REGION Network 17: STATE Num:30 StChkPalletPrsntL1L2
   RUNG wire#powerrail
      Contact( #s30_StChkPalletPrsntL1L2 )
      wire#w1
      I_Contact( #sStWtResetRel )
      I_Contact( #s30_StChkPalletPrsntL1L2_T1 )
      I_Contact( #s30_StChkPalletPrsntL1L2_T2 )
      I_Contact( #s30_StChkPalletPrsntL1L2_T3 )
      I_Contact( #s30_StChkPalletPrsntL1L2_T4 )
      wire#w2
      Coil( #s30_StChkPalletPrsntL1L2 )
   END_RUNG
   RUNG wire#powerrail
      Contact( #s20_StWtForL1L2StoprsUp_T1 )
   END_RUNG wire#w1
   RUNG wire#w2
      { S7_GenerateENO := "TRUE" } Move(in := 30, out1 => #StateNo)
   END_RUNG
   // the same network as SCL:
   #s30_StChkPalletPrsntL1L2 := (#s30_StChkPalletPrsntL1L2 OR #s20_StWtForL1L2StoprsUp_T1) AND NOT #sStWtResetRel AND NOT #s30_StChkPalletPrsntL1L2_T1 AND NOT #s30_StChkPalletPrsntL1L2_T2 AND NOT #s30_StChkPalletPrsntL1L2_T3 AND NOT #s30_StChkPalletPrsntL1L2_T4;
   IF #s30_StChkPalletPrsntL1L2 THEN #StateNo := 30; END_IF;
END_REGION

REGION Network 18: Transition for STATE Num:40 StChkPalletAtTT
   RUNG wire#powerrail
      Contact( #s40_StChkPalletAtTT )
      I_Contact( #sStWtResetRel )
      Contact( #sSst )
      wire#w1
      I_Contact( #iPalletAtTT )
      Coil( #s40_StChkPalletAtTT_T1 )
   END_RUNG
   RUNG wire#w1
      I_Contact( #s40_StChkPalletAtTT_T1 )
      Contact( #ipalletPrsntAtTT )
      Coil( #s40_StChkPalletAtTT_T2 )
   END_RUNG
   // the same network as SCL:
   #_w1 := #s40_StChkPalletAtTT AND NOT #sStWtResetRel AND #sSst;
   #s40_StChkPalletAtTT_T1 := #_w1 AND NOT #iPalletAtTT;
   #s40_StChkPalletAtTT_T2 := #_w1 AND NOT #s40_StChkPalletAtTT_T1 AND #ipalletPrsntAtTT;
END_REGION

REGION Network 19: STATE Num:40 StChkPalletAtTT
   RUNG wire#powerrail
      Contact( #s40_StChkPalletAtTT )
      wire#w1
      I_Contact( #sStWtResetRel )
      I_Contact( #s40_StChkPalletAtTT_T1 )
      I_Contact( #s40_StChkPalletAtTT_T2 )
      wire#w2
      Coil( #s40_StChkPalletAtTT )
   END_RUNG
   RUNG wire#powerrail
      Contact( #s30_StChkPalletPrsntL1L2_T1 )
   END_RUNG wire#w1
   RUNG wire#w2
      { S7_GenerateENO := "TRUE" } Move(in := 40, out1 => #StateNo)
   END_RUNG
   // the same network as SCL:
   #s40_StChkPalletAtTT := (#s40_StChkPalletAtTT OR #s30_StChkPalletPrsntL1L2_T1) AND NOT #sStWtResetRel AND NOT #s40_StChkPalletAtTT_T1 AND NOT #s40_StChkPalletAtTT_T2;
   IF #s40_StChkPalletAtTT THEN #StateNo := 40; END_IF;
END_REGION

REGION Network 20: Transition for STATE Num:50 StWtLifterAtPos1
   RUNG wire#powerrail
      Contact( #s50_StWtLifterAtPos1 )
      I_Contact( #sStWtResetRel )
      Contact( #sSst )
      Contact( #iLifterAtPos1 )
      Coil( #s50_StWtLifterAtPos1_T1 )
   END_RUNG
   // the same network as SCL:
   #s50_StWtLifterAtPos1_T1 := #s50_StWtLifterAtPos1 AND NOT #sStWtResetRel AND #sSst AND #iLifterAtPos1;
END_REGION

REGION Network 21: STATE Num:50 StWtLifterAtPos1
   RUNG wire#powerrail
      Contact( #s50_StWtLifterAtPos1 )
      wire#w1
      I_Contact( #sStWtResetRel )
      I_Contact( #s50_StWtLifterAtPos1_T1 )
      wire#w2
      Coil( #s50_StWtLifterAtPos1 )
   END_RUNG
   RUNG wire#powerrail
      Contact( #s40_StChkPalletAtTT_T1 )
   END_RUNG wire#w1
   RUNG wire#powerrail
      Contact( #s100_StRunOutActive_T1 )
   END_RUNG wire#w1
   RUNG wire#w2
      { S7_GenerateENO := "TRUE" } Move(in := 50, out1 => #StateNo)
   END_RUNG
   // the same network as SCL:
   #s50_StWtLifterAtPos1 := (#s50_StWtLifterAtPos1 OR #s40_StChkPalletAtTT_T1 OR #s100_StRunOutActive_T1) AND NOT #sStWtResetRel AND NOT #s50_StWtLifterAtPos1_T1;
   IF #s50_StWtLifterAtPos1 THEN #StateNo := 50; END_IF;
END_REGION

REGION Network 22: Actions for STATE Num:50 StWtLifterAtPos1
   RUNG wire#powerrail
      Contact( #s50_StWtLifterAtPos1 )
      Coil( #qLifterGotoPos1 )
   END_RUNG
   // the same network as SCL:
   #qLifterGotoPos1 := #s50_StWtLifterAtPos1;
END_REGION

REGION Network 23: Transition for STATE Num:60 StWtL1S2DownOver
   RUNG wire#powerrail
      Contact( #s60_StWtL1S2DownOver )
      I_Contact( #sStWtResetRel )
      Contact( #sSst )
      Contact( #iL1S2DownOver )
      Coil( #s60_StWtL1S2DownOver_T1 )
   END_RUNG
   // the same network as SCL:
   #s60_StWtL1S2DownOver_T1 := #s60_StWtL1S2DownOver AND NOT #sStWtResetRel AND #sSst AND #iL1S2DownOver;
END_REGION

REGION Network 24: STATE Num:60 StWtL1S2DownOver
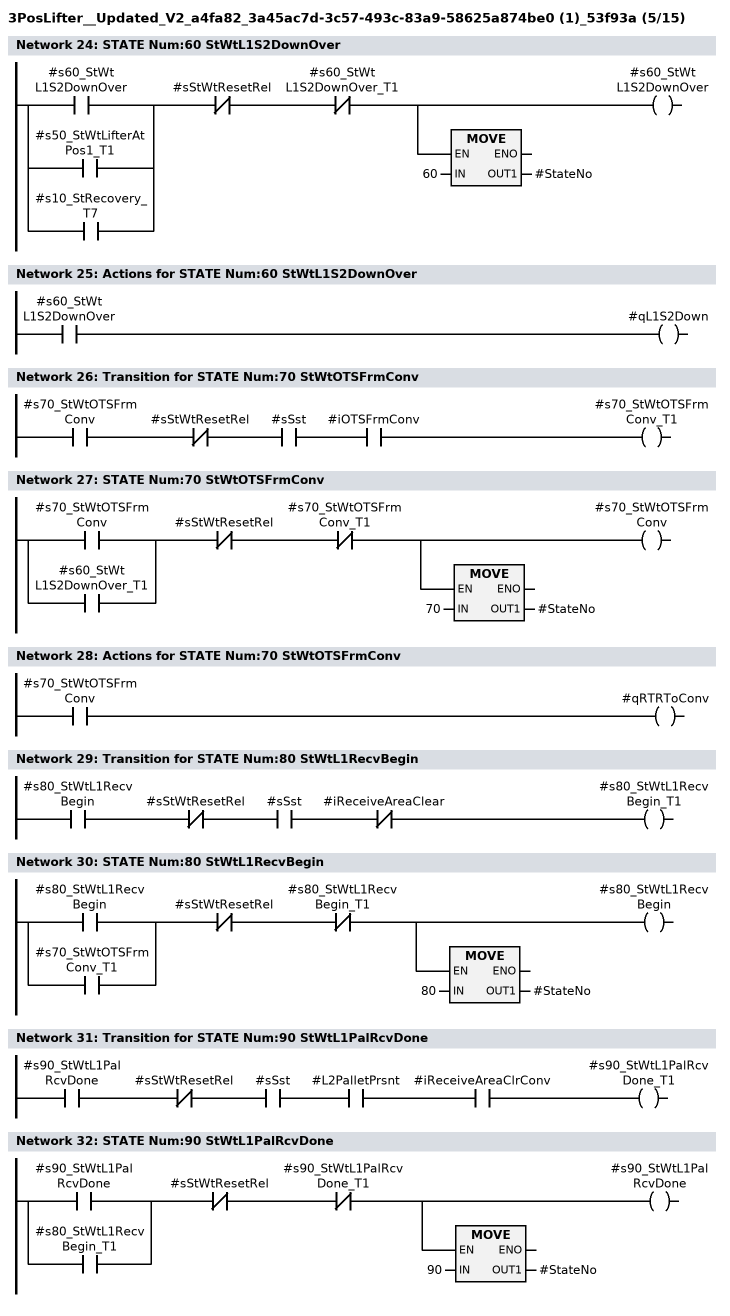
   RUNG wire#powerrail
      Contact( #s60_StWtL1S2DownOver )
      wire#w1
      I_Contact( #sStWtResetRel )
      I_Contact( #s60_StWtL1S2DownOver_T1 )
      wire#w2
      Coil( #s60_StWtL1S2DownOver )
   END_RUNG
   RUNG wire#powerrail
      Contact( #s50_StWtLifterAtPos1_T1 )
   END_RUNG wire#w1
   RUNG wire#powerrail
      Contact( #s10_StRecovery_T7 )
   END_RUNG wire#w1
   RUNG wire#w2
      { S7_GenerateENO := "TRUE" } Move(in := 60, out1 => #StateNo)
   END_RUNG
   // the same network as SCL:
   #s60_StWtL1S2DownOver := (#s60_StWtL1S2DownOver OR #s50_StWtLifterAtPos1_T1 OR #s10_StRecovery_T7) AND NOT #sStWtResetRel AND NOT #s60_StWtL1S2DownOver_T1;
   IF #s60_StWtL1S2DownOver THEN #StateNo := 60; END_IF;
END_REGION

REGION Network 25: Actions for STATE Num:60 StWtL1S2DownOver
   RUNG wire#powerrail
      Contact( #s60_StWtL1S2DownOver )
      Coil( #qL1S2Down )
   END_RUNG
   // the same network as SCL:
   #qL1S2Down := #s60_StWtL1S2DownOver;
END_REGION

REGION Network 26: Transition for STATE Num:70 StWtOTSFrmConv
   RUNG wire#powerrail
      Contact( #s70_StWtOTSFrmConv )
      I_Contact( #sStWtResetRel )
      Contact( #sSst )
      Contact( #iOTSFrmConv )
      Coil( #s70_StWtOTSFrmConv_T1 )
   END_RUNG
   // the same network as SCL:
   #s70_StWtOTSFrmConv_T1 := #s70_StWtOTSFrmConv AND NOT #sStWtResetRel AND #sSst AND #iOTSFrmConv;
END_REGION

REGION Network 27: STATE Num:70 StWtOTSFrmConv
   RUNG wire#powerrail
      Contact( #s70_StWtOTSFrmConv )
      wire#w1
      I_Contact( #sStWtResetRel )
      I_Contact( #s70_StWtOTSFrmConv_T1 )
      wire#w2
      Coil( #s70_StWtOTSFrmConv )
   END_RUNG
   RUNG wire#powerrail
      Contact( #s60_StWtL1S2DownOver_T1 )
   END_RUNG wire#w1
   RUNG wire#w2
      { S7_GenerateENO := "TRUE" } Move(in := 70, out1 => #StateNo)
   END_RUNG
   // the same network as SCL:
   #s70_StWtOTSFrmConv := (#s70_StWtOTSFrmConv OR #s60_StWtL1S2DownOver_T1) AND NOT #sStWtResetRel AND NOT #s70_StWtOTSFrmConv_T1;
   IF #s70_StWtOTSFrmConv THEN #StateNo := 70; END_IF;
END_REGION

REGION Network 28: Actions for STATE Num:70 StWtOTSFrmConv
   RUNG wire#powerrail
      Contact( #s70_StWtOTSFrmConv )
      Coil( #qRTRToConv )
   END_RUNG
   // the same network as SCL:
   #qRTRToConv := #s70_StWtOTSFrmConv;
END_REGION

REGION Network 29: Transition for STATE Num:80 StWtL1RecvBegin
   RUNG wire#powerrail
      Contact( #s80_StWtL1RecvBegin )
      I_Contact( #sStWtResetRel )
      Contact( #sSst )
      I_Contact( #iReceiveAreaClear )
      Coil( #s80_StWtL1RecvBegin_T1 )
   END_RUNG
   // the same network as SCL:
   #s80_StWtL1RecvBegin_T1 := #s80_StWtL1RecvBegin AND NOT #sStWtResetRel AND #sSst AND NOT #iReceiveAreaClear;
END_REGION

REGION Network 30: STATE Num:80 StWtL1RecvBegin
   RUNG wire#powerrail
      Contact( #s80_StWtL1RecvBegin )
      wire#w1
      I_Contact( #sStWtResetRel )
      I_Contact( #s80_StWtL1RecvBegin_T1 )
      wire#w2
      Coil( #s80_StWtL1RecvBegin )
   END_RUNG
   RUNG wire#powerrail
      Contact( #s70_StWtOTSFrmConv_T1 )
   END_RUNG wire#w1
   RUNG wire#w2
      { S7_GenerateENO := "TRUE" } Move(in := 80, out1 => #StateNo)
   END_RUNG
   // the same network as SCL:
   #s80_StWtL1RecvBegin := (#s80_StWtL1RecvBegin OR #s70_StWtOTSFrmConv_T1) AND NOT #sStWtResetRel AND NOT #s80_StWtL1RecvBegin_T1;
   IF #s80_StWtL1RecvBegin THEN #StateNo := 80; END_IF;
END_REGION

REGION Network 31: Transition for STATE Num:90 StWtL1PalRcvDone
   RUNG wire#powerrail
      Contact( #s90_StWtL1PalRcvDone )
      I_Contact( #sStWtResetRel )
      Contact( #sSst )
      Contact( #L2PalletPrsnt )
      Contact( #iReceiveAreaClrConv )
      Coil( #s90_StWtL1PalRcvDone_T1 )
   END_RUNG
   // the same network as SCL:
   #s90_StWtL1PalRcvDone_T1 := #s90_StWtL1PalRcvDone AND NOT #sStWtResetRel AND #sSst AND #L2PalletPrsnt AND #iReceiveAreaClrConv;
END_REGION

REGION Network 32: STATE Num:90 StWtL1PalRcvDone
   RUNG wire#powerrail
      Contact( #s90_StWtL1PalRcvDone )
      wire#w1
      I_Contact( #sStWtResetRel )
      I_Contact( #s90_StWtL1PalRcvDone_T1 )
      wire#w2
      Coil( #s90_StWtL1PalRcvDone )
   END_RUNG
   RUNG wire#powerrail
      Contact( #s80_StWtL1RecvBegin_T1 )
   END_RUNG wire#w1
   RUNG wire#w2
      { S7_GenerateENO := "TRUE" } Move(in := 90, out1 => #StateNo)
   END_RUNG
   // the same network as SCL:
   #s90_StWtL1PalRcvDone := (#s90_StWtL1PalRcvDone OR #s80_StWtL1RecvBegin_T1) AND NOT #sStWtResetRel AND NOT #s90_StWtL1PalRcvDone_T1;
   IF #s90_StWtL1PalRcvDone THEN #StateNo := 90; END_IF;
END_REGION

REGION Network 33: Transition for STATE Num:100 StRunOutActive
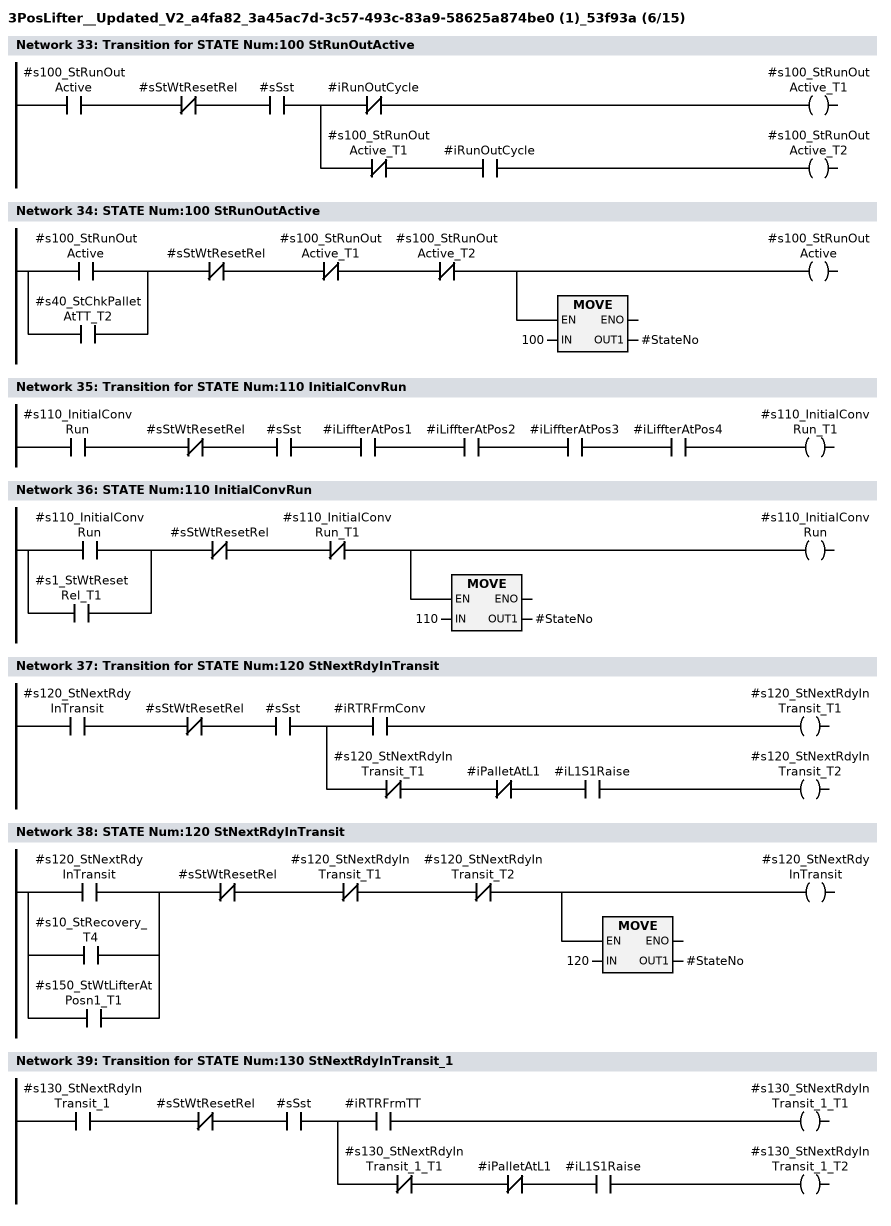
   RUNG wire#powerrail
      Contact( #s100_StRunOutActive )
      I_Contact( #sStWtResetRel )
      Contact( #sSst )
      wire#w1
      I_Contact( #iRunOutCycle )
      Coil( #s100_StRunOutActive_T1 )
   END_RUNG
   RUNG wire#w1
      I_Contact( #s100_StRunOutActive_T1 )
      Contact( #iRunOutCycle )
      Coil( #s100_StRunOutActive_T2 )
   END_RUNG
   // the same network as SCL:
   #_w1 := #s100_StRunOutActive AND NOT #sStWtResetRel AND #sSst;
   #s100_StRunOutActive_T1 := #_w1 AND NOT #iRunOutCycle;
   #s100_StRunOutActive_T2 := #_w1 AND NOT #s100_StRunOutActive_T1 AND #iRunOutCycle;
END_REGION

REGION Network 34: STATE Num:100 StRunOutActive
   RUNG wire#powerrail
      Contact( #s100_StRunOutActive )
      wire#w1
      I_Contact( #sStWtResetRel )
      I_Contact( #s100_StRunOutActive_T1 )
      I_Contact( #s100_StRunOutActive_T2 )
      wire#w2
      Coil( #s100_StRunOutActive )
   END_RUNG
   RUNG wire#powerrail
      Contact( #s40_StChkPalletAtTT_T2 )
   END_RUNG wire#w1
   RUNG wire#w2
      { S7_GenerateENO := "TRUE" } Move(in := 100, out1 => #StateNo)
   END_RUNG
   // the same network as SCL:
   #s100_StRunOutActive := (#s100_StRunOutActive OR #s40_StChkPalletAtTT_T2) AND NOT #sStWtResetRel AND NOT #s100_StRunOutActive_T1 AND NOT #s100_StRunOutActive_T2;
   IF #s100_StRunOutActive THEN #StateNo := 100; END_IF;
END_REGION

REGION Network 35: Transition for STATE Num:110 InitialConvRun
   RUNG wire#powerrail
      Contact( #s110_InitialConvRun )
      I_Contact( #sStWtResetRel )
      Contact( #sSst )
      Contact( #iLiffterAtPos1 )
      Contact( #iLiffterAtPos2 )
      Contact( #iLiffterAtPos3 )
      Contact( #iLiffterAtPos4 )
      Coil( #s110_InitialConvRun_T1 )
   END_RUNG
   // the same network as SCL:
   #s110_InitialConvRun_T1 := #s110_InitialConvRun AND NOT #sStWtResetRel AND #sSst AND #iLiffterAtPos1 AND #iLiffterAtPos2 AND #iLiffterAtPos3 AND #iLiffterAtPos4;
END_REGION

REGION Network 36: STATE Num:110 InitialConvRun
   RUNG wire#powerrail
      Contact( #s110_InitialConvRun )
      wire#w1
      I_Contact( #sStWtResetRel )
      I_Contact( #s110_InitialConvRun_T1 )
      wire#w2
      Coil( #s110_InitialConvRun )
   END_RUNG
   RUNG wire#powerrail
      Contact( #s1_StWtResetRel_T1 )
   END_RUNG wire#w1
   RUNG wire#w2
      { S7_GenerateENO := "TRUE" } Move(in := 110, out1 => #StateNo)
   END_RUNG
   // the same network as SCL:
   #s110_InitialConvRun := (#s110_InitialConvRun OR #s1_StWtResetRel_T1) AND NOT #sStWtResetRel AND NOT #s110_InitialConvRun_T1;
   IF #s110_InitialConvRun THEN #StateNo := 110; END_IF;
END_REGION

REGION Network 37: Transition for STATE Num:120 StNextRdyInTransit
   RUNG wire#powerrail
      Contact( #s120_StNextRdyInTransit )
      I_Contact( #sStWtResetRel )
      Contact( #sSst )
      wire#w1
      Contact( #iRTRFrmConv )
      Coil( #s120_StNextRdyInTransit_T1 )
   END_RUNG
   RUNG wire#w1
      I_Contact( #s120_StNextRdyInTransit_T1 )
      I_Contact( #iPalletAtL1 )
      Contact( #iL1S1Raise )
      Coil( #s120_StNextRdyInTransit_T2 )
   END_RUNG
   // the same network as SCL:
   #_w1 := #s120_StNextRdyInTransit AND NOT #sStWtResetRel AND #sSst;
   #s120_StNextRdyInTransit_T1 := #_w1 AND #iRTRFrmConv;
   #s120_StNextRdyInTransit_T2 := #_w1 AND NOT #s120_StNextRdyInTransit_T1 AND NOT #iPalletAtL1 AND #iL1S1Raise;
END_REGION

REGION Network 38: STATE Num:120 StNextRdyInTransit
   RUNG wire#powerrail
      Contact( #s120_StNextRdyInTransit )
      wire#w1
      I_Contact( #sStWtResetRel )
      I_Contact( #s120_StNextRdyInTransit_T1 )
      I_Contact( #s120_StNextRdyInTransit_T2 )
      wire#w2
      Coil( #s120_StNextRdyInTransit )
   END_RUNG
   RUNG wire#powerrail
      Contact( #s10_StRecovery_T4 )
   END_RUNG wire#w1
   RUNG wire#powerrail
      Contact( #s150_StWtLifterAtPosn1_T1 )
   END_RUNG wire#w1
   RUNG wire#w2
      { S7_GenerateENO := "TRUE" } Move(in := 120, out1 => #StateNo)
   END_RUNG
   // the same network as SCL:
   #s120_StNextRdyInTransit := (#s120_StNextRdyInTransit OR #s10_StRecovery_T4 OR #s150_StWtLifterAtPosn1_T1) AND NOT #sStWtResetRel AND NOT #s120_StNextRdyInTransit_T1 AND NOT #s120_StNextRdyInTransit_T2;
   IF #s120_StNextRdyInTransit THEN #StateNo := 120; END_IF;
END_REGION

REGION Network 39: Transition for STATE Num:130 StNextRdyInTransit_1
   RUNG wire#powerrail
      Contact( #s130_StNextRdyInTransit_1 )
      I_Contact( #sStWtResetRel )
      Contact( #sSst )
      wire#w1
      Contact( #iRTRFrmTT )
      Coil( #s130_StNextRdyInTransit_1_T1 )
   END_RUNG
   RUNG wire#w1
      I_Contact( #s130_StNextRdyInTransit_1_T1 )
      I_Contact( #iPalletAtL1 )
      Contact( #iL1S1Raise )
      Coil( #s130_StNextRdyInTransit_1_T2 )
   END_RUNG
   // the same network as SCL:
   #_w1 := #s130_StNextRdyInTransit_1 AND NOT #sStWtResetRel AND #sSst;
   #s130_StNextRdyInTransit_1_T1 := #_w1 AND #iRTRFrmTT;
   #s130_StNextRdyInTransit_1_T2 := #_w1 AND NOT #s130_StNextRdyInTransit_1_T1 AND NOT #iPalletAtL1 AND #iL1S1Raise;
END_REGION

REGION Network 40: STATE Num:130 StNextRdyInTransit_1
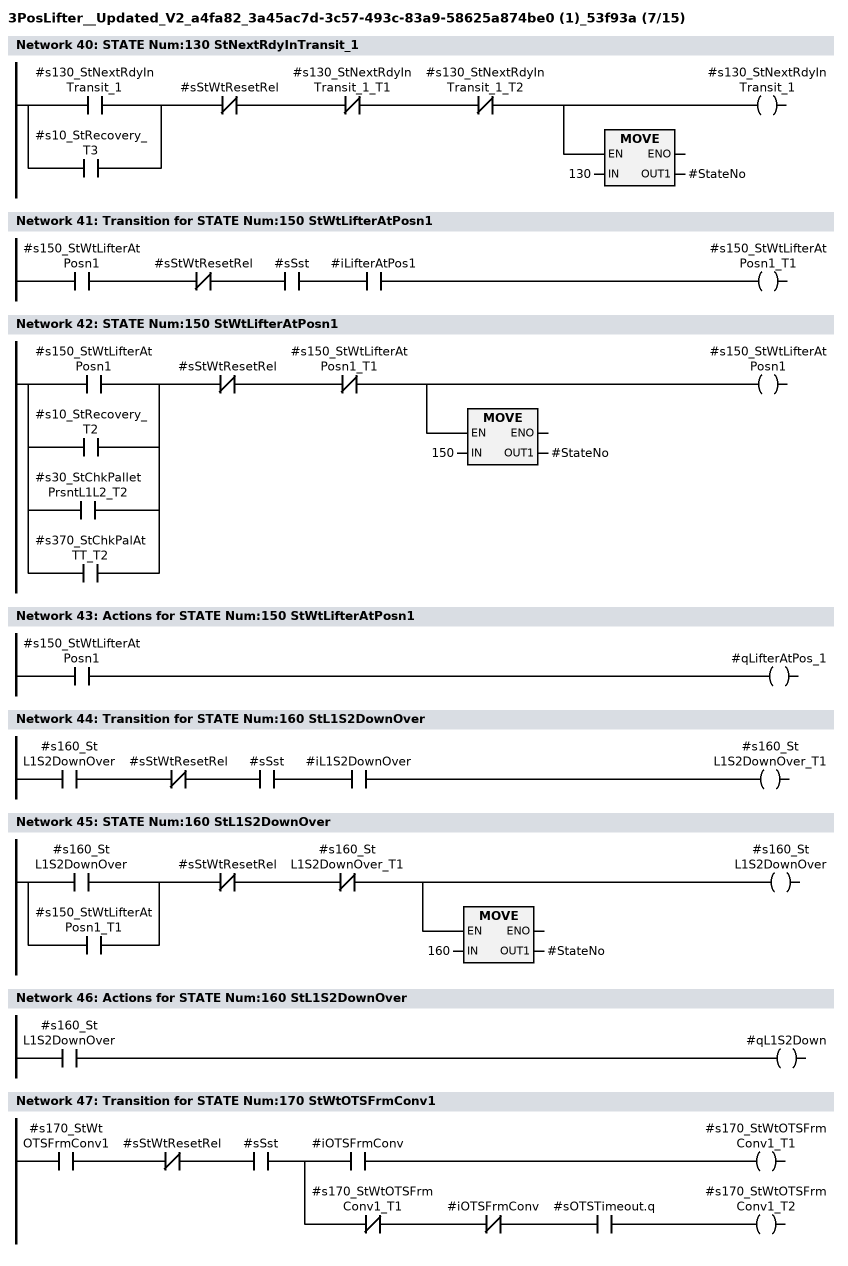
   RUNG wire#powerrail
      Contact( #s130_StNextRdyInTransit_1 )
      wire#w1
      I_Contact( #sStWtResetRel )
      I_Contact( #s130_StNextRdyInTransit_1_T1 )
      I_Contact( #s130_StNextRdyInTransit_1_T2 )
      wire#w2
      Coil( #s130_StNextRdyInTransit_1 )
   END_RUNG
   RUNG wire#powerrail
      Contact( #s10_StRecovery_T3 )
   END_RUNG wire#w1
   RUNG wire#w2
      { S7_GenerateENO := "TRUE" } Move(in := 130, out1 => #StateNo)
   END_RUNG
   // the same network as SCL:
   #s130_StNextRdyInTransit_1 := (#s130_StNextRdyInTransit_1 OR #s10_StRecovery_T3) AND NOT #sStWtResetRel AND NOT #s130_StNextRdyInTransit_1_T1 AND NOT #s130_StNextRdyInTransit_1_T2;
   IF #s130_StNextRdyInTransit_1 THEN #StateNo := 130; END_IF;
END_REGION

REGION Network 41: Transition for STATE Num:150 StWtLifterAtPosn1
   RUNG wire#powerrail
      Contact( #s150_StWtLifterAtPosn1 )
      I_Contact( #sStWtResetRel )
      Contact( #sSst )
      Contact( #iLifterAtPos1 )
      Coil( #s150_StWtLifterAtPosn1_T1 )
   END_RUNG
   // the same network as SCL:
   #s150_StWtLifterAtPosn1_T1 := #s150_StWtLifterAtPosn1 AND NOT #sStWtResetRel AND #sSst AND #iLifterAtPos1;
END_REGION

REGION Network 42: STATE Num:150 StWtLifterAtPosn1
   RUNG wire#powerrail
      Contact( #s150_StWtLifterAtPosn1 )
      wire#w1
      I_Contact( #sStWtResetRel )
      I_Contact( #s150_StWtLifterAtPosn1_T1 )
      wire#w2
      Coil( #s150_StWtLifterAtPosn1 )
   END_RUNG
   RUNG wire#powerrail
      Contact( #s10_StRecovery_T2 )
   END_RUNG wire#w1
   RUNG wire#powerrail
      Contact( #s30_StChkPalletPrsntL1L2_T2 )
   END_RUNG wire#w1
   RUNG wire#powerrail
      Contact( #s370_StChkPalAtTT_T2 )
   END_RUNG wire#w1
   RUNG wire#w2
      { S7_GenerateENO := "TRUE" } Move(in := 150, out1 => #StateNo)
   END_RUNG
   // the same network as SCL:
   #s150_StWtLifterAtPosn1 := (#s150_StWtLifterAtPosn1 OR #s10_StRecovery_T2 OR #s30_StChkPalletPrsntL1L2_T2 OR #s370_StChkPalAtTT_T2) AND NOT #sStWtResetRel AND NOT #s150_StWtLifterAtPosn1_T1;
   IF #s150_StWtLifterAtPosn1 THEN #StateNo := 150; END_IF;
END_REGION

REGION Network 43: Actions for STATE Num:150 StWtLifterAtPosn1
   RUNG wire#powerrail
      Contact( #s150_StWtLifterAtPosn1 )
      Coil( #qLifterAtPos_1 )
   END_RUNG
   // the same network as SCL:
   #qLifterAtPos_1 := #s150_StWtLifterAtPosn1;
END_REGION

REGION Network 44: Transition for STATE Num:160 StL1S2DownOver
   RUNG wire#powerrail
      Contact( #s160_StL1S2DownOver )
      I_Contact( #sStWtResetRel )
      Contact( #sSst )
      Contact( #iL1S2DownOver )
      Coil( #s160_StL1S2DownOver_T1 )
   END_RUNG
   // the same network as SCL:
   #s160_StL1S2DownOver_T1 := #s160_StL1S2DownOver AND NOT #sStWtResetRel AND #sSst AND #iL1S2DownOver;
END_REGION

REGION Network 45: STATE Num:160 StL1S2DownOver
   RUNG wire#powerrail
      Contact( #s160_StL1S2DownOver )
      wire#w1
      I_Contact( #sStWtResetRel )
      I_Contact( #s160_StL1S2DownOver_T1 )
      wire#w2
      Coil( #s160_StL1S2DownOver )
   END_RUNG
   RUNG wire#powerrail
      Contact( #s150_StWtLifterAtPosn1_T1 )
   END_RUNG wire#w1
   RUNG wire#w2
      { S7_GenerateENO := "TRUE" } Move(in := 160, out1 => #StateNo)
   END_RUNG
   // the same network as SCL:
   #s160_StL1S2DownOver := (#s160_StL1S2DownOver OR #s150_StWtLifterAtPosn1_T1) AND NOT #sStWtResetRel AND NOT #s160_StL1S2DownOver_T1;
   IF #s160_StL1S2DownOver THEN #StateNo := 160; END_IF;
END_REGION

REGION Network 46: Actions for STATE Num:160 StL1S2DownOver
   RUNG wire#powerrail
      Contact( #s160_StL1S2DownOver )
      Coil( #qL1S2Down )
   END_RUNG
   // the same network as SCL:
   #qL1S2Down := #s160_StL1S2DownOver;
END_REGION

REGION Network 47: Transition for STATE Num:170 StWtOTSFrmConv1
   RUNG wire#powerrail
      Contact( #s170_StWtOTSFrmConv1 )
      I_Contact( #sStWtResetRel )
      Contact( #sSst )
      wire#w1
      Contact( #iOTSFrmConv )
      Coil( #s170_StWtOTSFrmConv1_T1 )
   END_RUNG
   RUNG wire#w1
      I_Contact( #s170_StWtOTSFrmConv1_T1 )
      I_Contact( #iOTSFrmConv )
      Contact( #sOTSTimeout.q )
      Coil( #s170_StWtOTSFrmConv1_T2 )
   END_RUNG
   // the same network as SCL:
   #_w1 := #s170_StWtOTSFrmConv1 AND NOT #sStWtResetRel AND #sSst;
   #s170_StWtOTSFrmConv1_T1 := #_w1 AND #iOTSFrmConv;
   #s170_StWtOTSFrmConv1_T2 := #_w1 AND NOT #s170_StWtOTSFrmConv1_T1 AND NOT #iOTSFrmConv AND #sOTSTimeout.q;
END_REGION

REGION Network 48: STATE Num:170 StWtOTSFrmConv1
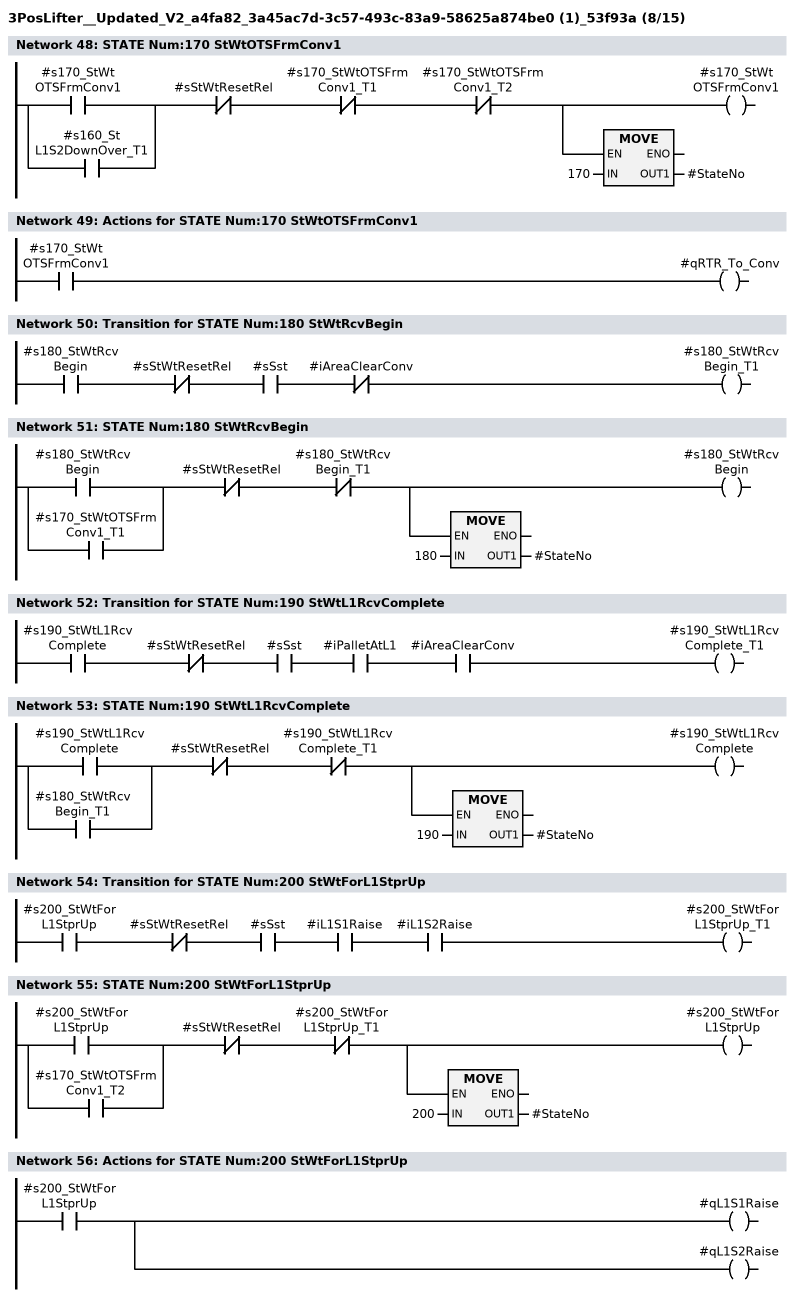
   RUNG wire#powerrail
      Contact( #s170_StWtOTSFrmConv1 )
      wire#w1
      I_Contact( #sStWtResetRel )
      I_Contact( #s170_StWtOTSFrmConv1_T1 )
      I_Contact( #s170_StWtOTSFrmConv1_T2 )
      wire#w2
      Coil( #s170_StWtOTSFrmConv1 )
   END_RUNG
   RUNG wire#powerrail
      Contact( #s160_StL1S2DownOver_T1 )
   END_RUNG wire#w1
   RUNG wire#w2
      { S7_GenerateENO := "TRUE" } Move(in := 170, out1 => #StateNo)
   END_RUNG
   // the same network as SCL:
   #s170_StWtOTSFrmConv1 := (#s170_StWtOTSFrmConv1 OR #s160_StL1S2DownOver_T1) AND NOT #sStWtResetRel AND NOT #s170_StWtOTSFrmConv1_T1 AND NOT #s170_StWtOTSFrmConv1_T2;
   IF #s170_StWtOTSFrmConv1 THEN #StateNo := 170; END_IF;
END_REGION

REGION Network 49: Actions for STATE Num:170 StWtOTSFrmConv1
   RUNG wire#powerrail
      Contact( #s170_StWtOTSFrmConv1 )
      Coil( #qRTR_To_Conv )
   END_RUNG
   // the same network as SCL:
   #qRTR_To_Conv := #s170_StWtOTSFrmConv1;
END_REGION

REGION Network 50: Transition for STATE Num:180 StWtRcvBegin
   RUNG wire#powerrail
      Contact( #s180_StWtRcvBegin )
      I_Contact( #sStWtResetRel )
      Contact( #sSst )
      I_Contact( #iAreaClearConv )
      Coil( #s180_StWtRcvBegin_T1 )
   END_RUNG
   // the same network as SCL:
   #s180_StWtRcvBegin_T1 := #s180_StWtRcvBegin AND NOT #sStWtResetRel AND #sSst AND NOT #iAreaClearConv;
END_REGION

REGION Network 51: STATE Num:180 StWtRcvBegin
   RUNG wire#powerrail
      Contact( #s180_StWtRcvBegin )
      wire#w1
      I_Contact( #sStWtResetRel )
      I_Contact( #s180_StWtRcvBegin_T1 )
      wire#w2
      Coil( #s180_StWtRcvBegin )
   END_RUNG
   RUNG wire#powerrail
      Contact( #s170_StWtOTSFrmConv1_T1 )
   END_RUNG wire#w1
   RUNG wire#w2
      { S7_GenerateENO := "TRUE" } Move(in := 180, out1 => #StateNo)
   END_RUNG
   // the same network as SCL:
   #s180_StWtRcvBegin := (#s180_StWtRcvBegin OR #s170_StWtOTSFrmConv1_T1) AND NOT #sStWtResetRel AND NOT #s180_StWtRcvBegin_T1;
   IF #s180_StWtRcvBegin THEN #StateNo := 180; END_IF;
END_REGION

REGION Network 52: Transition for STATE Num:190 StWtL1RcvComplete
   RUNG wire#powerrail
      Contact( #s190_StWtL1RcvComplete )
      I_Contact( #sStWtResetRel )
      Contact( #sSst )
      Contact( #iPalletAtL1 )
      Contact( #iAreaClearConv )
      Coil( #s190_StWtL1RcvComplete_T1 )
   END_RUNG
   // the same network as SCL:
   #s190_StWtL1RcvComplete_T1 := #s190_StWtL1RcvComplete AND NOT #sStWtResetRel AND #sSst AND #iPalletAtL1 AND #iAreaClearConv;
END_REGION

REGION Network 53: STATE Num:190 StWtL1RcvComplete
   RUNG wire#powerrail
      Contact( #s190_StWtL1RcvComplete )
      wire#w1
      I_Contact( #sStWtResetRel )
      I_Contact( #s190_StWtL1RcvComplete_T1 )
      wire#w2
      Coil( #s190_StWtL1RcvComplete )
   END_RUNG
   RUNG wire#powerrail
      Contact( #s180_StWtRcvBegin_T1 )
   END_RUNG wire#w1
   RUNG wire#w2
      { S7_GenerateENO := "TRUE" } Move(in := 190, out1 => #StateNo)
   END_RUNG
   // the same network as SCL:
   #s190_StWtL1RcvComplete := (#s190_StWtL1RcvComplete OR #s180_StWtRcvBegin_T1) AND NOT #sStWtResetRel AND NOT #s190_StWtL1RcvComplete_T1;
   IF #s190_StWtL1RcvComplete THEN #StateNo := 190; END_IF;
END_REGION

REGION Network 54: Transition for STATE Num:200 StWtForL1StprUp
   RUNG wire#powerrail
      Contact( #s200_StWtForL1StprUp )
      I_Contact( #sStWtResetRel )
      Contact( #sSst )
      Contact( #iL1S1Raise )
      Contact( #iL1S2Raise )
      Coil( #s200_StWtForL1StprUp_T1 )
   END_RUNG
   // the same network as SCL:
   #s200_StWtForL1StprUp_T1 := #s200_StWtForL1StprUp AND NOT #sStWtResetRel AND #sSst AND #iL1S1Raise AND #iL1S2Raise;
END_REGION

REGION Network 55: STATE Num:200 StWtForL1StprUp
   RUNG wire#powerrail
      Contact( #s200_StWtForL1StprUp )
      wire#w1
      I_Contact( #sStWtResetRel )
      I_Contact( #s200_StWtForL1StprUp_T1 )
      wire#w2
      Coil( #s200_StWtForL1StprUp )
   END_RUNG
   RUNG wire#powerrail
      Contact( #s170_StWtOTSFrmConv1_T2 )
   END_RUNG wire#w1
   RUNG wire#w2
      { S7_GenerateENO := "TRUE" } Move(in := 200, out1 => #StateNo)
   END_RUNG
   // the same network as SCL:
   #s200_StWtForL1StprUp := (#s200_StWtForL1StprUp OR #s170_StWtOTSFrmConv1_T2) AND NOT #sStWtResetRel AND NOT #s200_StWtForL1StprUp_T1;
   IF #s200_StWtForL1StprUp THEN #StateNo := 200; END_IF;
END_REGION

REGION Network 56: Actions for STATE Num:200 StWtForL1StprUp
   RUNG wire#powerrail
      Contact( #s200_StWtForL1StprUp )
      wire#w1
      Coil( #qL1S1Raise )
   END_RUNG
   RUNG wire#w1
      Coil( #qL1S2Raise )
   END_RUNG
   // the same network as SCL:
   #qL1S1Raise := #s200_StWtForL1StprUp;
   #qL1S2Raise := #s200_StWtForL1StprUp;
END_REGION

REGION Network 57: Transition for STATE Num:220 StWtL2S2Down
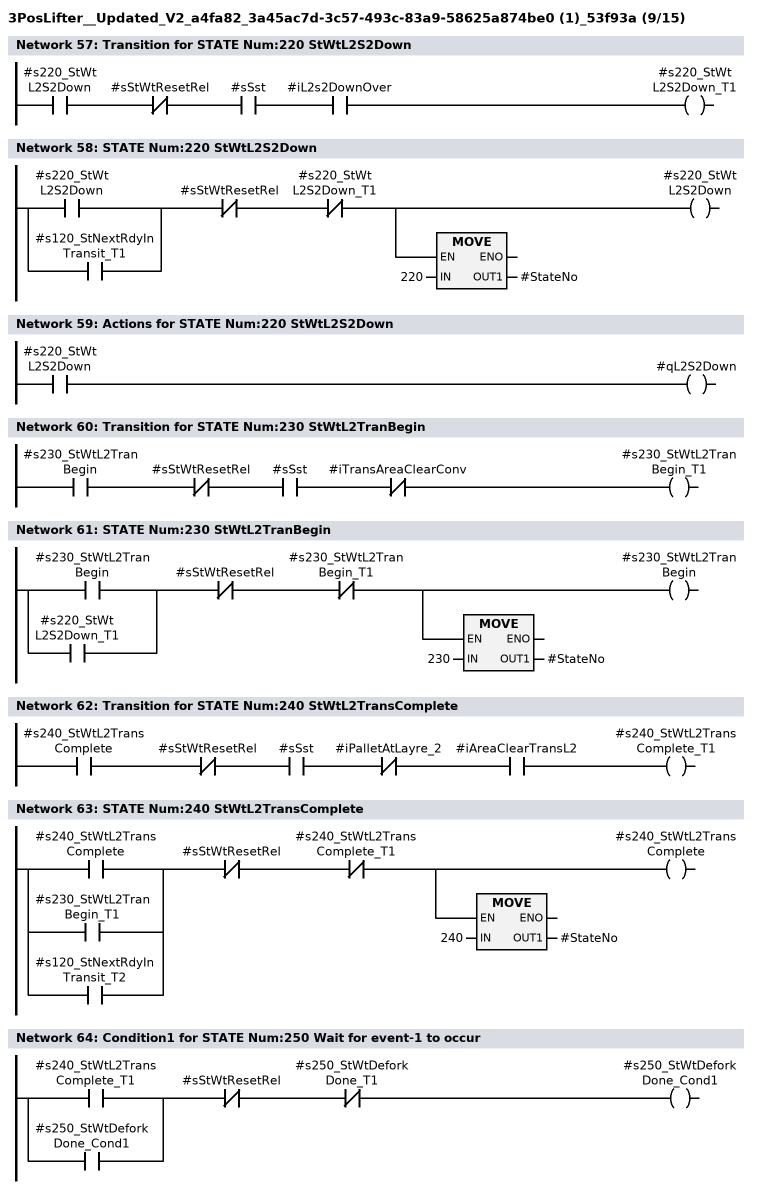
   RUNG wire#powerrail
      Contact( #s220_StWtL2S2Down )
      I_Contact( #sStWtResetRel )
      Contact( #sSst )
      Contact( #iL2s2DownOver )
      Coil( #s220_StWtL2S2Down_T1 )
   END_RUNG
   // the same network as SCL:
   #s220_StWtL2S2Down_T1 := #s220_StWtL2S2Down AND NOT #sStWtResetRel AND #sSst AND #iL2s2DownOver;
END_REGION

REGION Network 58: STATE Num:220 StWtL2S2Down
   RUNG wire#powerrail
      Contact( #s220_StWtL2S2Down )
      wire#w1
      I_Contact( #sStWtResetRel )
      I_Contact( #s220_StWtL2S2Down_T1 )
      wire#w2
      Coil( #s220_StWtL2S2Down )
   END_RUNG
   RUNG wire#powerrail
      Contact( #s120_StNextRdyInTransit_T1 )
   END_RUNG wire#w1
   RUNG wire#w2
      { S7_GenerateENO := "TRUE" } Move(in := 220, out1 => #StateNo)
   END_RUNG
   // the same network as SCL:
   #s220_StWtL2S2Down := (#s220_StWtL2S2Down OR #s120_StNextRdyInTransit_T1) AND NOT #sStWtResetRel AND NOT #s220_StWtL2S2Down_T1;
   IF #s220_StWtL2S2Down THEN #StateNo := 220; END_IF;
END_REGION

REGION Network 59: Actions for STATE Num:220 StWtL2S2Down
   RUNG wire#powerrail
      Contact( #s220_StWtL2S2Down )
      Coil( #qL2S2Down )
   END_RUNG
   // the same network as SCL:
   #qL2S2Down := #s220_StWtL2S2Down;
END_REGION

REGION Network 60: Transition for STATE Num:230 StWtL2TranBegin
   RUNG wire#powerrail
      Contact( #s230_StWtL2TranBegin )
      I_Contact( #sStWtResetRel )
      Contact( #sSst )
      I_Contact( #iTransAreaClearConv )
      Coil( #s230_StWtL2TranBegin_T1 )
   END_RUNG
   // the same network as SCL:
   #s230_StWtL2TranBegin_T1 := #s230_StWtL2TranBegin AND NOT #sStWtResetRel AND #sSst AND NOT #iTransAreaClearConv;
END_REGION

REGION Network 61: STATE Num:230 StWtL2TranBegin
   RUNG wire#powerrail
      Contact( #s230_StWtL2TranBegin )
      wire#w1
      I_Contact( #sStWtResetRel )
      I_Contact( #s230_StWtL2TranBegin_T1 )
      wire#w2
      Coil( #s230_StWtL2TranBegin )
   END_RUNG
   RUNG wire#powerrail
      Contact( #s220_StWtL2S2Down_T1 )
   END_RUNG wire#w1
   RUNG wire#w2
      { S7_GenerateENO := "TRUE" } Move(in := 230, out1 => #StateNo)
   END_RUNG
   // the same network as SCL:
   #s230_StWtL2TranBegin := (#s230_StWtL2TranBegin OR #s220_StWtL2S2Down_T1) AND NOT #sStWtResetRel AND NOT #s230_StWtL2TranBegin_T1;
   IF #s230_StWtL2TranBegin THEN #StateNo := 230; END_IF;
END_REGION

REGION Network 62: Transition for STATE Num:240 StWtL2TransComplete
   RUNG wire#powerrail
      Contact( #s240_StWtL2TransComplete )
      I_Contact( #sStWtResetRel )
      Contact( #sSst )
      I_Contact( #iPalletAtLayre_2 )
      Contact( #iAreaClearTransL2 )
      Coil( #s240_StWtL2TransComplete_T1 )
   END_RUNG
   // the same network as SCL:
   #s240_StWtL2TransComplete_T1 := #s240_StWtL2TransComplete AND NOT #sStWtResetRel AND #sSst AND NOT #iPalletAtLayre_2 AND #iAreaClearTransL2;
END_REGION

REGION Network 63: STATE Num:240 StWtL2TransComplete
   RUNG wire#powerrail
      Contact( #s240_StWtL2TransComplete )
      wire#w1
      I_Contact( #sStWtResetRel )
      I_Contact( #s240_StWtL2TransComplete_T1 )
      wire#w2
      Coil( #s240_StWtL2TransComplete )
   END_RUNG
   RUNG wire#powerrail
      Contact( #s230_StWtL2TranBegin_T1 )
   END_RUNG wire#w1
   RUNG wire#powerrail
      Contact( #s120_StNextRdyInTransit_T2 )
   END_RUNG wire#w1
   RUNG wire#w2
      { S7_GenerateENO := "TRUE" } Move(in := 240, out1 => #StateNo)
   END_RUNG
   // the same network as SCL:
   #s240_StWtL2TransComplete := (#s240_StWtL2TransComplete OR #s230_StWtL2TranBegin_T1 OR #s120_StNextRdyInTransit_T2) AND NOT #sStWtResetRel AND NOT #s240_StWtL2TransComplete_T1;
   IF #s240_StWtL2TransComplete THEN #StateNo := 240; END_IF;
END_REGION

REGION Network 64: Condition1 for STATE Num:250 Wait for event-1 to occur
   RUNG wire#powerrail
      Contact( #s240_StWtL2TransComplete_T1 )
      wire#w1
      I_Contact( #sStWtResetRel )
      I_Contact( #s250_StWtDeforkDone_T1 )
      Coil( #s250_StWtDeforkDone_Cond1 )
   END_RUNG
   RUNG wire#powerrail
      Contact( #s250_StWtDeforkDone_Cond1 )
   END_RUNG wire#w1
   // the same network as SCL:
   #s250_StWtDeforkDone_Cond1 := (#s240_StWtL2TransComplete_T1 OR #s250_StWtDeforkDone_Cond1) AND NOT #sStWtResetRel AND NOT #s250_StWtDeforkDone_T1;
END_REGION

REGION Network 65: Condition2 for STATE Num:250 Wait for event-1 to occur
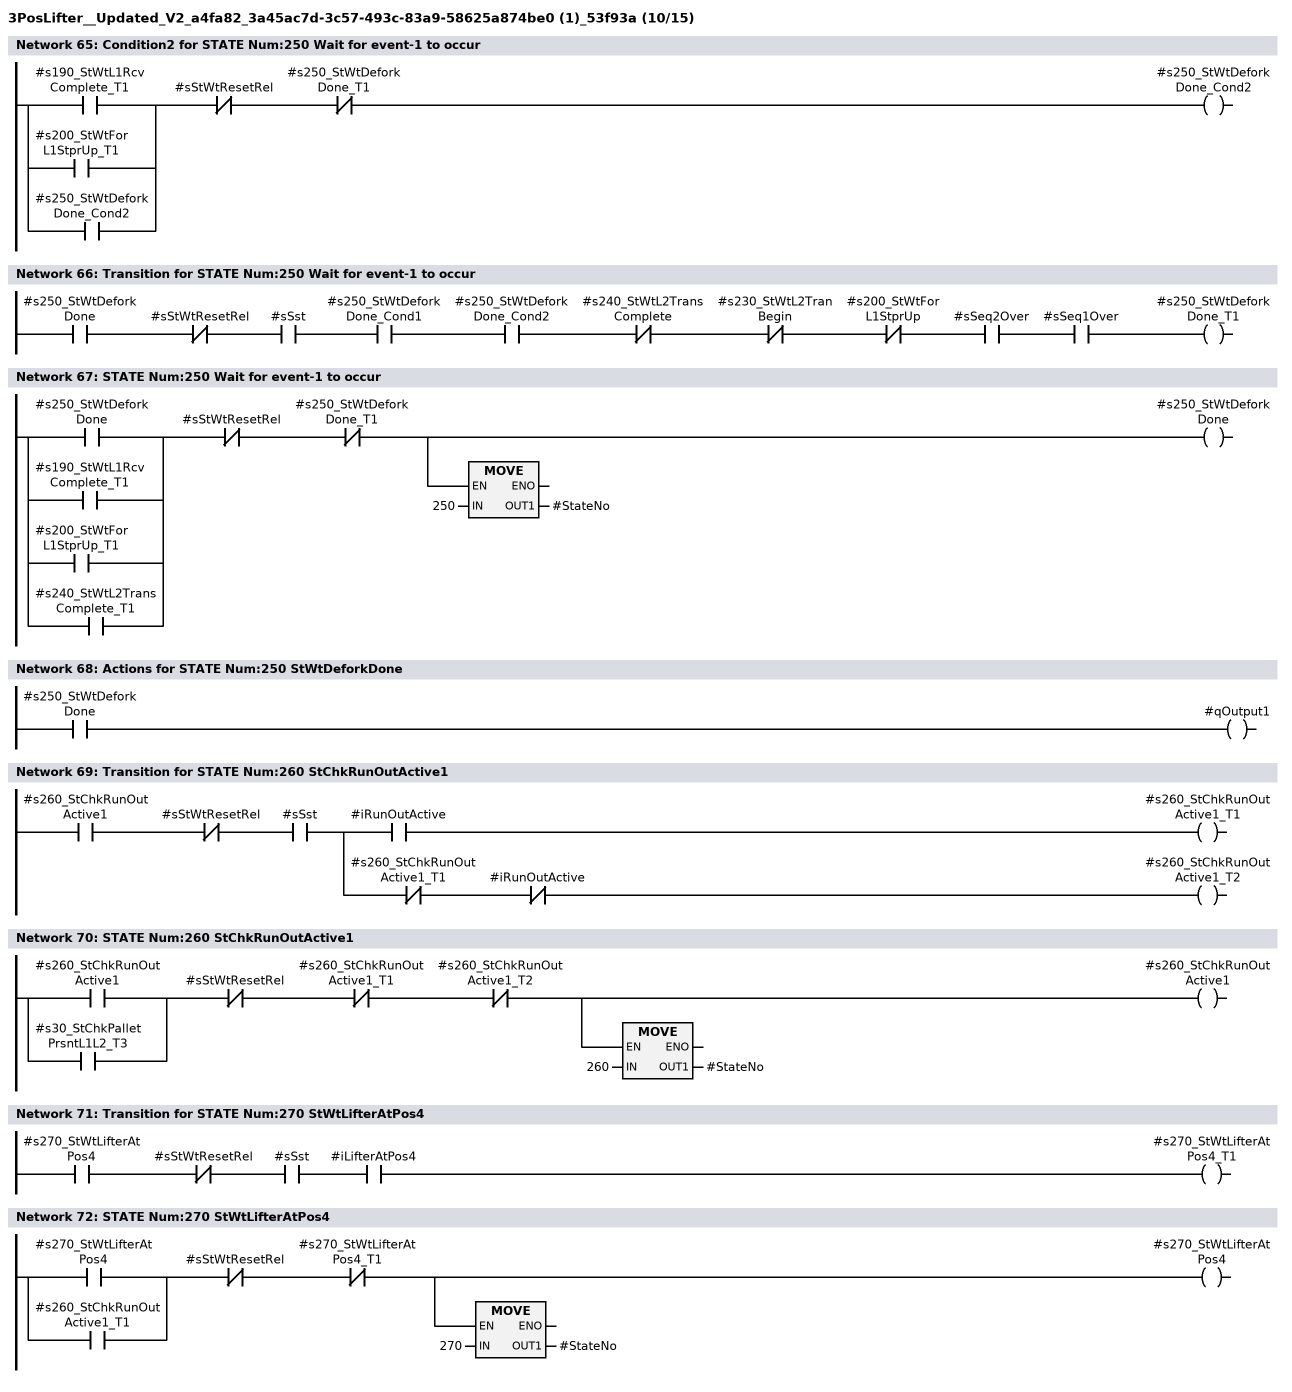
   RUNG wire#powerrail
      Contact( #s190_StWtL1RcvComplete_T1 )
      wire#w1
      I_Contact( #sStWtResetRel )
      I_Contact( #s250_StWtDeforkDone_T1 )
      Coil( #s250_StWtDeforkDone_Cond2 )
   END_RUNG
   RUNG wire#powerrail
      Contact( #s200_StWtForL1StprUp_T1 )
   END_RUNG wire#w1
   RUNG wire#powerrail
      Contact( #s250_StWtDeforkDone_Cond2 )
   END_RUNG wire#w1
   // the same network as SCL:
   #s250_StWtDeforkDone_Cond2 := (#s190_StWtL1RcvComplete_T1 OR #s200_StWtForL1StprUp_T1 OR #s250_StWtDeforkDone_Cond2) AND NOT #sStWtResetRel AND NOT #s250_StWtDeforkDone_T1;
END_REGION

REGION Network 66: Transition for STATE Num:250 Wait for event-1 to occur
   RUNG wire#powerrail
      Contact( #s250_StWtDeforkDone )
      I_Contact( #sStWtResetRel )
      Contact( #sSst )
      Contact( #s250_StWtDeforkDone_Cond1 )
      Contact( #s250_StWtDeforkDone_Cond2 )
      I_Contact( #s240_StWtL2TransComplete )
      I_Contact( #s230_StWtL2TranBegin )
      I_Contact( #s200_StWtForL1StprUp )
      Contact( #sSeq2Over )
      Contact( #sSeq1Over )
      Coil( #s250_StWtDeforkDone_T1 )
   END_RUNG
   // the same network as SCL:
   #s250_StWtDeforkDone_T1 := #s250_StWtDeforkDone AND NOT #sStWtResetRel AND #sSst AND #s250_StWtDeforkDone_Cond1 AND #s250_StWtDeforkDone_Cond2 AND NOT #s240_StWtL2TransComplete AND NOT #s230_StWtL2TranBegin AND NOT #s200_StWtForL1StprUp AND #sSeq2Over AND #sSeq1Over;
END_REGION

REGION Network 67: STATE Num:250 Wait for event-1 to occur
   RUNG wire#powerrail
      Contact( #s250_StWtDeforkDone )
      wire#w1
      I_Contact( #sStWtResetRel )
      I_Contact( #s250_StWtDeforkDone_T1 )
      wire#w2
      Coil( #s250_StWtDeforkDone )
   END_RUNG
   RUNG wire#powerrail
      Contact( #s190_StWtL1RcvComplete_T1 )
   END_RUNG wire#w1
   RUNG wire#powerrail
      Contact( #s200_StWtForL1StprUp_T1 )
   END_RUNG wire#w1
   RUNG wire#powerrail
      Contact( #s240_StWtL2TransComplete_T1 )
   END_RUNG wire#w1
   RUNG wire#w2
      { S7_GenerateENO := "TRUE" } Move(in := 250, out1 => #StateNo)
   END_RUNG
   // the same network as SCL:
   #s250_StWtDeforkDone := (#s250_StWtDeforkDone OR #s190_StWtL1RcvComplete_T1 OR #s200_StWtForL1StprUp_T1 OR #s240_StWtL2TransComplete_T1) AND NOT #sStWtResetRel AND NOT #s250_StWtDeforkDone_T1;
   IF #s250_StWtDeforkDone THEN #StateNo := 250; END_IF;
END_REGION

REGION Network 68: Actions for STATE Num:250 StWtDeforkDone
   RUNG wire#powerrail
      Contact( #s250_StWtDeforkDone )
      Coil( #qOutput1 )
   END_RUNG
   // the same network as SCL:
   #qOutput1 := #s250_StWtDeforkDone;
END_REGION

REGION Network 69: Transition for STATE Num:260 StChkRunOutActive1
   RUNG wire#powerrail
      Contact( #s260_StChkRunOutActive1 )
      I_Contact( #sStWtResetRel )
      Contact( #sSst )
      wire#w1
      Contact( #iRunOutActive )
      Coil( #s260_StChkRunOutActive1_T1 )
   END_RUNG
   RUNG wire#w1
      I_Contact( #s260_StChkRunOutActive1_T1 )
      I_Contact( #iRunOutActive )
      Coil( #s260_StChkRunOutActive1_T2 )
   END_RUNG
   // the same network as SCL:
   #_w1 := #s260_StChkRunOutActive1 AND NOT #sStWtResetRel AND #sSst;
   #s260_StChkRunOutActive1_T1 := #_w1 AND #iRunOutActive;
   #s260_StChkRunOutActive1_T2 := #_w1 AND NOT #s260_StChkRunOutActive1_T1 AND NOT #iRunOutActive;
END_REGION

REGION Network 70: STATE Num:260 StChkRunOutActive1
   RUNG wire#powerrail
      Contact( #s260_StChkRunOutActive1 )
      wire#w1
      I_Contact( #sStWtResetRel )
      I_Contact( #s260_StChkRunOutActive1_T1 )
      I_Contact( #s260_StChkRunOutActive1_T2 )
      wire#w2
      Coil( #s260_StChkRunOutActive1 )
   END_RUNG
   RUNG wire#powerrail
      Contact( #s30_StChkPalletPrsntL1L2_T3 )
   END_RUNG wire#w1
   RUNG wire#w2
      { S7_GenerateENO := "TRUE" } Move(in := 260, out1 => #StateNo)
   END_RUNG
   // the same network as SCL:
   #s260_StChkRunOutActive1 := (#s260_StChkRunOutActive1 OR #s30_StChkPalletPrsntL1L2_T3) AND NOT #sStWtResetRel AND NOT #s260_StChkRunOutActive1_T1 AND NOT #s260_StChkRunOutActive1_T2;
   IF #s260_StChkRunOutActive1 THEN #StateNo := 260; END_IF;
END_REGION

REGION Network 71: Transition for STATE Num:270 StWtLifterAtPos4
   RUNG wire#powerrail
      Contact( #s270_StWtLifterAtPos4 )
      I_Contact( #sStWtResetRel )
      Contact( #sSst )
      Contact( #iLifterAtPos4 )
      Coil( #s270_StWtLifterAtPos4_T1 )
   END_RUNG
   // the same network as SCL:
   #s270_StWtLifterAtPos4_T1 := #s270_StWtLifterAtPos4 AND NOT #sStWtResetRel AND #sSst AND #iLifterAtPos4;
END_REGION

REGION Network 72: STATE Num:270 StWtLifterAtPos4
   RUNG wire#powerrail
      Contact( #s270_StWtLifterAtPos4 )
      wire#w1
      I_Contact( #sStWtResetRel )
      I_Contact( #s270_StWtLifterAtPos4_T1 )
      wire#w2
      Coil( #s270_StWtLifterAtPos4 )
   END_RUNG
   RUNG wire#powerrail
      Contact( #s260_StChkRunOutActive1_T1 )
   END_RUNG wire#w1
   RUNG wire#w2
      { S7_GenerateENO := "TRUE" } Move(in := 270, out1 => #StateNo)
   END_RUNG
   // the same network as SCL:
   #s270_StWtLifterAtPos4 := (#s270_StWtLifterAtPos4 OR #s260_StChkRunOutActive1_T1) AND NOT #sStWtResetRel AND NOT #s270_StWtLifterAtPos4_T1;
   IF #s270_StWtLifterAtPos4 THEN #StateNo := 270; END_IF;
END_REGION

REGION Network 73: Actions for STATE Num:270 StWtLifterAtPos4
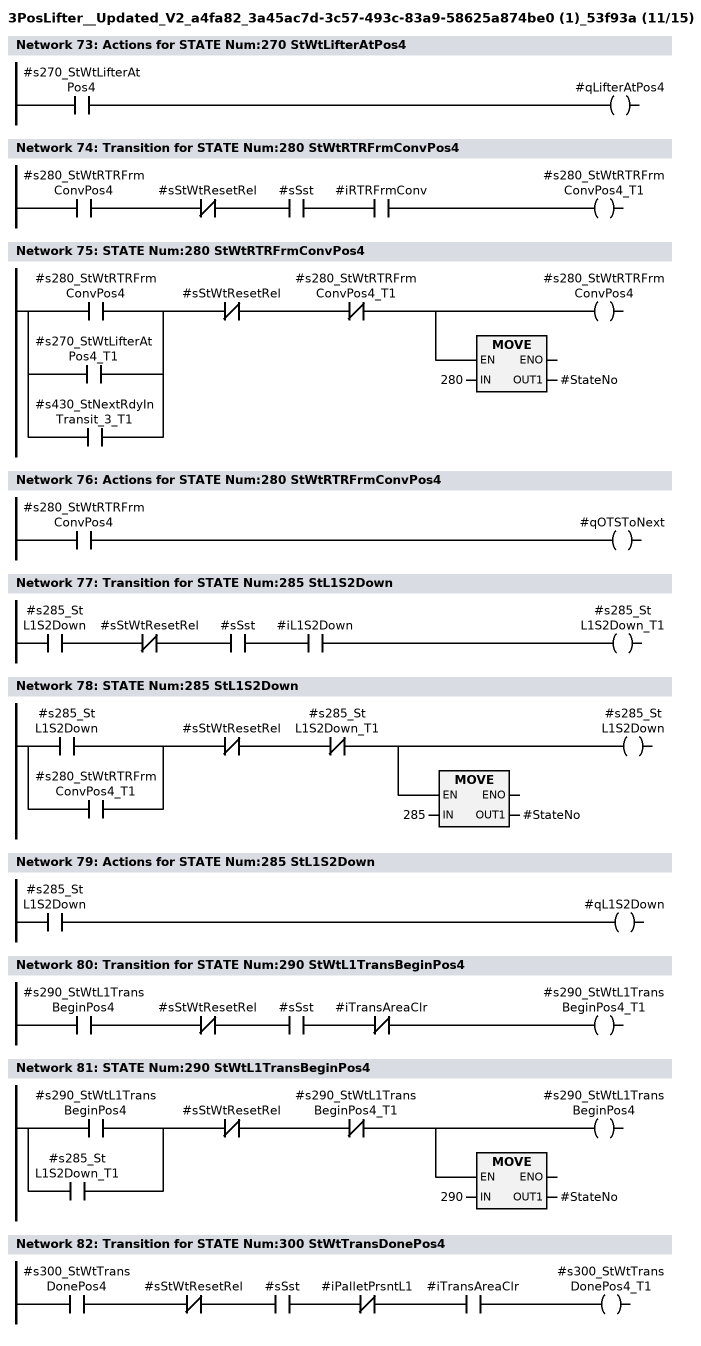
   RUNG wire#powerrail
      Contact( #s270_StWtLifterAtPos4 )
      Coil( #qLifterAtPos4 )
   END_RUNG
   // the same network as SCL:
   #qLifterAtPos4 := #s270_StWtLifterAtPos4;
END_REGION

REGION Network 74: Transition for STATE Num:280 StWtRTRFrmConvPos4
   RUNG wire#powerrail
      Contact( #s280_StWtRTRFrmConvPos4 )
      I_Contact( #sStWtResetRel )
      Contact( #sSst )
      Contact( #iRTRFrmConv )
      Coil( #s280_StWtRTRFrmConvPos4_T1 )
   END_RUNG
   // the same network as SCL:
   #s280_StWtRTRFrmConvPos4_T1 := #s280_StWtRTRFrmConvPos4 AND NOT #sStWtResetRel AND #sSst AND #iRTRFrmConv;
END_REGION

REGION Network 75: STATE Num:280 StWtRTRFrmConvPos4
   RUNG wire#powerrail
      Contact( #s280_StWtRTRFrmConvPos4 )
      wire#w1
      I_Contact( #sStWtResetRel )
      I_Contact( #s280_StWtRTRFrmConvPos4_T1 )
      wire#w2
      Coil( #s280_StWtRTRFrmConvPos4 )
   END_RUNG
   RUNG wire#powerrail
      Contact( #s270_StWtLifterAtPos4_T1 )
   END_RUNG wire#w1
   RUNG wire#powerrail
      Contact( #s430_StNextRdyInTransit_3_T1 )
   END_RUNG wire#w1
   RUNG wire#w2
      { S7_GenerateENO := "TRUE" } Move(in := 280, out1 => #StateNo)
   END_RUNG
   // the same network as SCL:
   #s280_StWtRTRFrmConvPos4 := (#s280_StWtRTRFrmConvPos4 OR #s270_StWtLifterAtPos4_T1 OR #s430_StNextRdyInTransit_3_T1) AND NOT #sStWtResetRel AND NOT #s280_StWtRTRFrmConvPos4_T1;
   IF #s280_StWtRTRFrmConvPos4 THEN #StateNo := 280; END_IF;
END_REGION

REGION Network 76: Actions for STATE Num:280 StWtRTRFrmConvPos4
   RUNG wire#powerrail
      Contact( #s280_StWtRTRFrmConvPos4 )
      Coil( #qOTSToNext )
   END_RUNG
   // the same network as SCL:
   #qOTSToNext := #s280_StWtRTRFrmConvPos4;
END_REGION

REGION Network 77: Transition for STATE Num:285 StL1S2Down
   RUNG wire#powerrail
      Contact( #s285_StL1S2Down )
      I_Contact( #sStWtResetRel )
      Contact( #sSst )
      Contact( #iL1S2Down )
      Coil( #s285_StL1S2Down_T1 )
   END_RUNG
   // the same network as SCL:
   #s285_StL1S2Down_T1 := #s285_StL1S2Down AND NOT #sStWtResetRel AND #sSst AND #iL1S2Down;
END_REGION

REGION Network 78: STATE Num:285 StL1S2Down
   RUNG wire#powerrail
      Contact( #s285_StL1S2Down )
      wire#w1
      I_Contact( #sStWtResetRel )
      I_Contact( #s285_StL1S2Down_T1 )
      wire#w2
      Coil( #s285_StL1S2Down )
   END_RUNG
   RUNG wire#powerrail
      Contact( #s280_StWtRTRFrmConvPos4_T1 )
   END_RUNG wire#w1
   RUNG wire#w2
      { S7_GenerateENO := "TRUE" } Move(in := 285, out1 => #StateNo)
   END_RUNG
   // the same network as SCL:
   #s285_StL1S2Down := (#s285_StL1S2Down OR #s280_StWtRTRFrmConvPos4_T1) AND NOT #sStWtResetRel AND NOT #s285_StL1S2Down_T1;
   IF #s285_StL1S2Down THEN #StateNo := 285; END_IF;
END_REGION

REGION Network 79: Actions for STATE Num:285 StL1S2Down
   RUNG wire#powerrail
      Contact( #s285_StL1S2Down )
      Coil( #qL1S2Down )
   END_RUNG
   // the same network as SCL:
   #qL1S2Down := #s285_StL1S2Down;
END_REGION

REGION Network 80: Transition for STATE Num:290 StWtL1TransBeginPos4
   RUNG wire#powerrail
      Contact( #s290_StWtL1TransBeginPos4 )
      I_Contact( #sStWtResetRel )
      Contact( #sSst )
      I_Contact( #iTransAreaClr )
      Coil( #s290_StWtL1TransBeginPos4_T1 )
   END_RUNG
   // the same network as SCL:
   #s290_StWtL1TransBeginPos4_T1 := #s290_StWtL1TransBeginPos4 AND NOT #sStWtResetRel AND #sSst AND NOT #iTransAreaClr;
END_REGION

REGION Network 81: STATE Num:290 StWtL1TransBeginPos4
   RUNG wire#powerrail
      Contact( #s290_StWtL1TransBeginPos4 )
      wire#w1
      I_Contact( #sStWtResetRel )
      I_Contact( #s290_StWtL1TransBeginPos4_T1 )
      wire#w2
      Coil( #s290_StWtL1TransBeginPos4 )
   END_RUNG
   RUNG wire#powerrail
      Contact( #s285_StL1S2Down_T1 )
   END_RUNG wire#w1
   RUNG wire#w2
      { S7_GenerateENO := "TRUE" } Move(in := 290, out1 => #StateNo)
   END_RUNG
   // the same network as SCL:
   #s290_StWtL1TransBeginPos4 := (#s290_StWtL1TransBeginPos4 OR #s285_StL1S2Down_T1) AND NOT #sStWtResetRel AND NOT #s290_StWtL1TransBeginPos4_T1;
   IF #s290_StWtL1TransBeginPos4 THEN #StateNo := 290; END_IF;
END_REGION

REGION Network 82: Transition for STATE Num:300 StWtTransDonePos4
   RUNG wire#powerrail
      Contact( #s300_StWtTransDonePos4 )
      I_Contact( #sStWtResetRel )
      Contact( #sSst )
      I_Contact( #iPalletPrsntL1 )
      Contact( #iTransAreaClr )
      Coil( #s300_StWtTransDonePos4_T1 )
   END_RUNG
   // the same network as SCL:
   #s300_StWtTransDonePos4_T1 := #s300_StWtTransDonePos4 AND NOT #sStWtResetRel AND #sSst AND NOT #iPalletPrsntL1 AND #iTransAreaClr;
END_REGION

REGION Network 83: STATE Num:300 StWtTransDonePos4
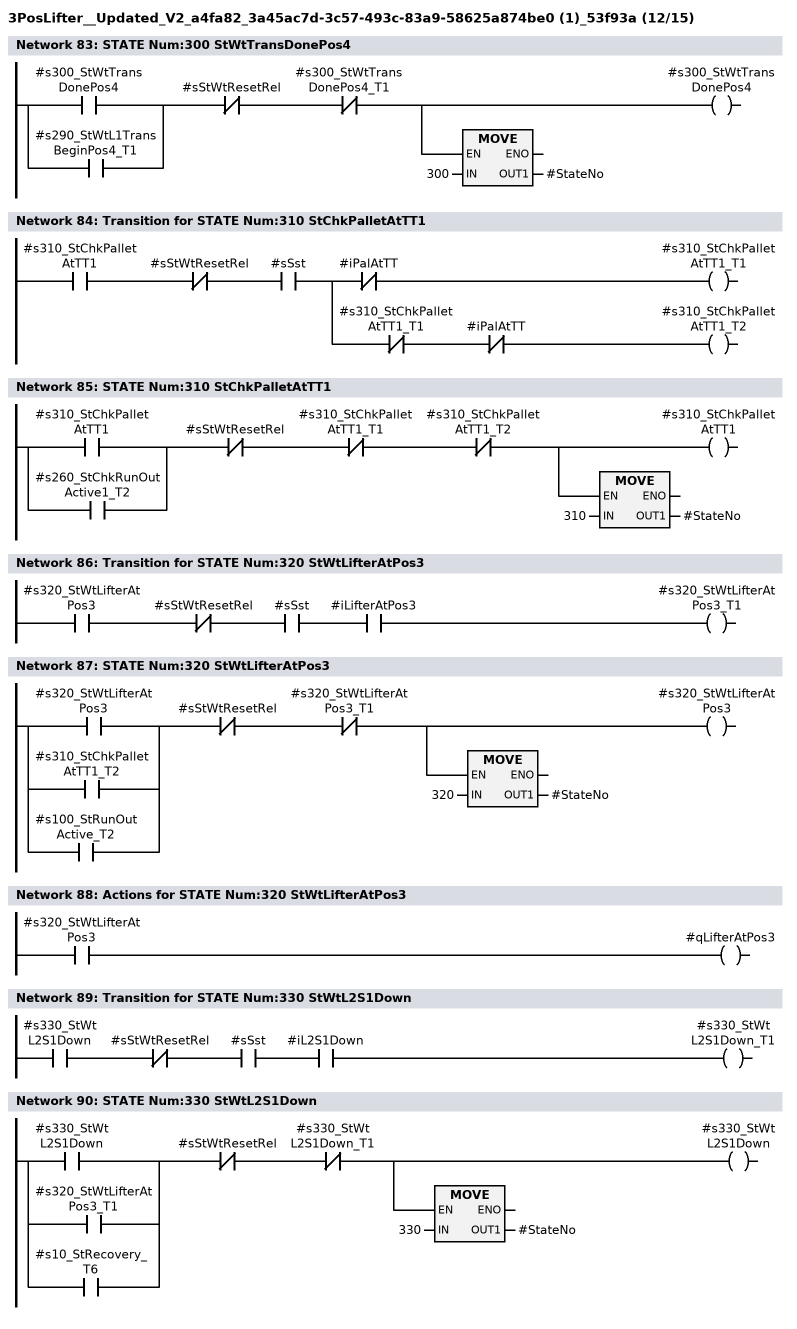
   RUNG wire#powerrail
      Contact( #s300_StWtTransDonePos4 )
      wire#w1
      I_Contact( #sStWtResetRel )
      I_Contact( #s300_StWtTransDonePos4_T1 )
      wire#w2
      Coil( #s300_StWtTransDonePos4 )
   END_RUNG
   RUNG wire#powerrail
      Contact( #s290_StWtL1TransBeginPos4_T1 )
   END_RUNG wire#w1
   RUNG wire#w2
      { S7_GenerateENO := "TRUE" } Move(in := 300, out1 => #StateNo)
   END_RUNG
   // the same network as SCL:
   #s300_StWtTransDonePos4 := (#s300_StWtTransDonePos4 OR #s290_StWtL1TransBeginPos4_T1) AND NOT #sStWtResetRel AND NOT #s300_StWtTransDonePos4_T1;
   IF #s300_StWtTransDonePos4 THEN #StateNo := 300; END_IF;
END_REGION

REGION Network 84: Transition for STATE Num:310 StChkPalletAtTT1
   RUNG wire#powerrail
      Contact( #s310_StChkPalletAtTT1 )
      I_Contact( #sStWtResetRel )
      Contact( #sSst )
      wire#w1
      I_Contact( #iPalAtTT )
      Coil( #s310_StChkPalletAtTT1_T1 )
   END_RUNG
   RUNG wire#w1
      I_Contact( #s310_StChkPalletAtTT1_T1 )
      I_Contact( #iPalAtTT )
      Coil( #s310_StChkPalletAtTT1_T2 )
   END_RUNG
   // the same network as SCL:
   #_w1 := #s310_StChkPalletAtTT1 AND NOT #sStWtResetRel AND #sSst;
   #s310_StChkPalletAtTT1_T1 := #_w1 AND NOT #iPalAtTT;
   #s310_StChkPalletAtTT1_T2 := #_w1 AND NOT #s310_StChkPalletAtTT1_T1 AND NOT #iPalAtTT;
END_REGION

REGION Network 85: STATE Num:310 StChkPalletAtTT1
   RUNG wire#powerrail
      Contact( #s310_StChkPalletAtTT1 )
      wire#w1
      I_Contact( #sStWtResetRel )
      I_Contact( #s310_StChkPalletAtTT1_T1 )
      I_Contact( #s310_StChkPalletAtTT1_T2 )
      wire#w2
      Coil( #s310_StChkPalletAtTT1 )
   END_RUNG
   RUNG wire#powerrail
      Contact( #s260_StChkRunOutActive1_T2 )
   END_RUNG wire#w1
   RUNG wire#w2
      { S7_GenerateENO := "TRUE" } Move(in := 310, out1 => #StateNo)
   END_RUNG
   // the same network as SCL:
   #s310_StChkPalletAtTT1 := (#s310_StChkPalletAtTT1 OR #s260_StChkRunOutActive1_T2) AND NOT #sStWtResetRel AND NOT #s310_StChkPalletAtTT1_T1 AND NOT #s310_StChkPalletAtTT1_T2;
   IF #s310_StChkPalletAtTT1 THEN #StateNo := 310; END_IF;
END_REGION

REGION Network 86: Transition for STATE Num:320 StWtLifterAtPos3
   RUNG wire#powerrail
      Contact( #s320_StWtLifterAtPos3 )
      I_Contact( #sStWtResetRel )
      Contact( #sSst )
      Contact( #iLifterAtPos3 )
      Coil( #s320_StWtLifterAtPos3_T1 )
   END_RUNG
   // the same network as SCL:
   #s320_StWtLifterAtPos3_T1 := #s320_StWtLifterAtPos3 AND NOT #sStWtResetRel AND #sSst AND #iLifterAtPos3;
END_REGION

REGION Network 87: STATE Num:320 StWtLifterAtPos3
   RUNG wire#powerrail
      Contact( #s320_StWtLifterAtPos3 )
      wire#w1
      I_Contact( #sStWtResetRel )
      I_Contact( #s320_StWtLifterAtPos3_T1 )
      wire#w2
      Coil( #s320_StWtLifterAtPos3 )
   END_RUNG
   RUNG wire#powerrail
      Contact( #s310_StChkPalletAtTT1_T2 )
   END_RUNG wire#w1
   RUNG wire#powerrail
      Contact( #s100_StRunOutActive_T2 )
   END_RUNG wire#w1
   RUNG wire#w2
      { S7_GenerateENO := "TRUE" } Move(in := 320, out1 => #StateNo)
   END_RUNG
   // the same network as SCL:
   #s320_StWtLifterAtPos3 := (#s320_StWtLifterAtPos3 OR #s310_StChkPalletAtTT1_T2 OR #s100_StRunOutActive_T2) AND NOT #sStWtResetRel AND NOT #s320_StWtLifterAtPos3_T1;
   IF #s320_StWtLifterAtPos3 THEN #StateNo := 320; END_IF;
END_REGION

REGION Network 88: Actions for STATE Num:320 StWtLifterAtPos3
   RUNG wire#powerrail
      Contact( #s320_StWtLifterAtPos3 )
      Coil( #qLifterAtPos3 )
   END_RUNG
   // the same network as SCL:
   #qLifterAtPos3 := #s320_StWtLifterAtPos3;
END_REGION

REGION Network 89: Transition for STATE Num:330 StWtL2S1Down
   RUNG wire#powerrail
      Contact( #s330_StWtL2S1Down )
      I_Contact( #sStWtResetRel )
      Contact( #sSst )
      Contact( #iL2S1Down )
      Coil( #s330_StWtL2S1Down_T1 )
   END_RUNG
   // the same network as SCL:
   #s330_StWtL2S1Down_T1 := #s330_StWtL2S1Down AND NOT #sStWtResetRel AND #sSst AND #iL2S1Down;
END_REGION

REGION Network 90: STATE Num:330 StWtL2S1Down
   RUNG wire#powerrail
      Contact( #s330_StWtL2S1Down )
      wire#w1
      I_Contact( #sStWtResetRel )
      I_Contact( #s330_StWtL2S1Down_T1 )
      wire#w2
      Coil( #s330_StWtL2S1Down )
   END_RUNG
   RUNG wire#powerrail
      Contact( #s320_StWtLifterAtPos3_T1 )
   END_RUNG wire#w1
   RUNG wire#powerrail
      Contact( #s10_StRecovery_T6 )
   END_RUNG wire#w1
   RUNG wire#w2
      { S7_GenerateENO := "TRUE" } Move(in := 330, out1 => #StateNo)
   END_RUNG
   // the same network as SCL:
   #s330_StWtL2S1Down := (#s330_StWtL2S1Down OR #s320_StWtLifterAtPos3_T1 OR #s10_StRecovery_T6) AND NOT #sStWtResetRel AND NOT #s330_StWtL2S1Down_T1;
   IF #s330_StWtL2S1Down THEN #StateNo := 330; END_IF;
END_REGION

REGION Network 91: Actions for STATE Num:330 StWtL2S1Down
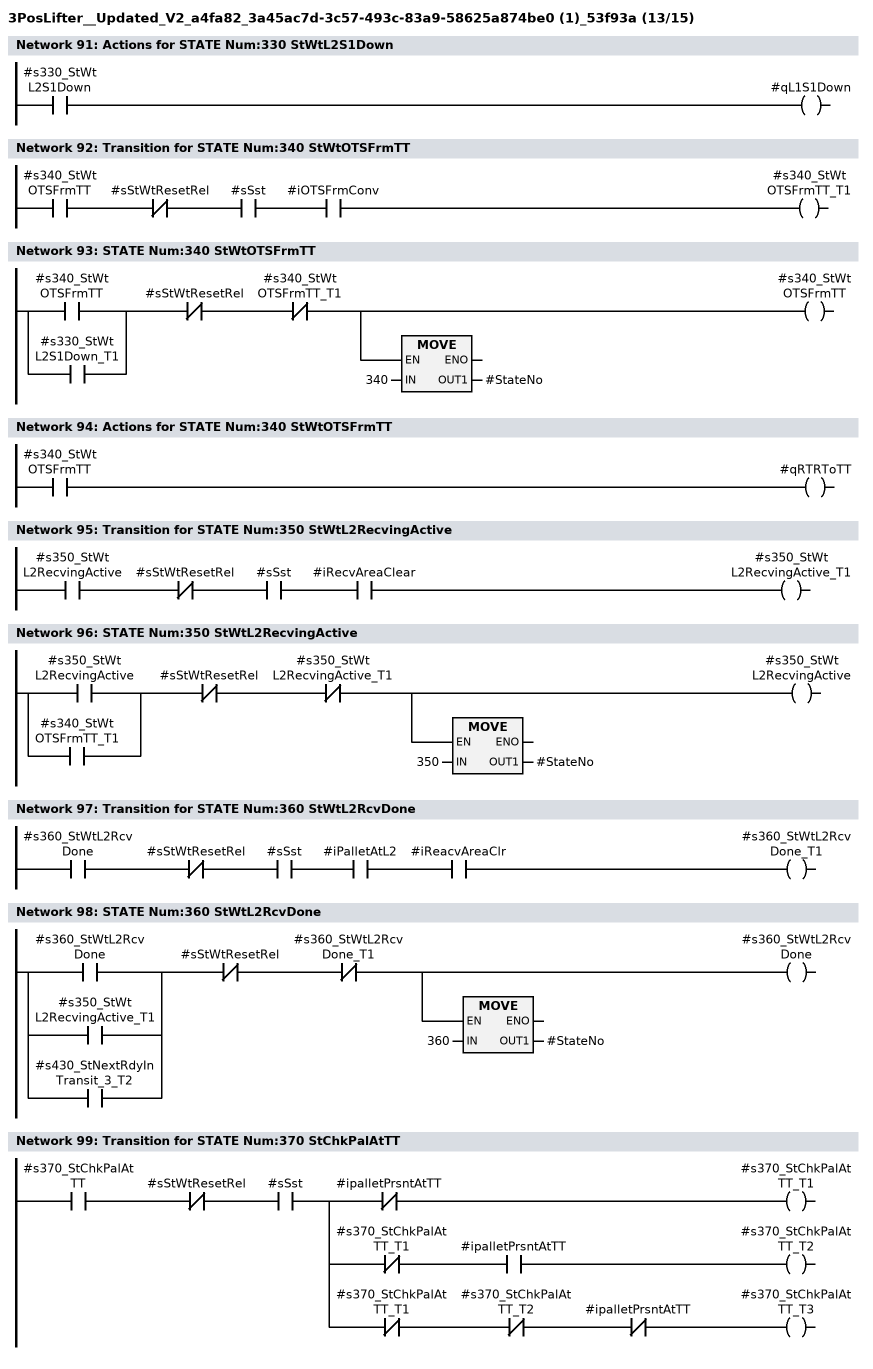
   RUNG wire#powerrail
      Contact( #s330_StWtL2S1Down )
      Coil( #qL1S1Down )
   END_RUNG
   // the same network as SCL:
   #qL1S1Down := #s330_StWtL2S1Down;
END_REGION

REGION Network 92: Transition for STATE Num:340 StWtOTSFrmTT
   RUNG wire#powerrail
      Contact( #s340_StWtOTSFrmTT )
      I_Contact( #sStWtResetRel )
      Contact( #sSst )
      Contact( #iOTSFrmConv )
      Coil( #s340_StWtOTSFrmTT_T1 )
   END_RUNG
   // the same network as SCL:
   #s340_StWtOTSFrmTT_T1 := #s340_StWtOTSFrmTT AND NOT #sStWtResetRel AND #sSst AND #iOTSFrmConv;
END_REGION

REGION Network 93: STATE Num:340 StWtOTSFrmTT
   RUNG wire#powerrail
      Contact( #s340_StWtOTSFrmTT )
      wire#w1
      I_Contact( #sStWtResetRel )
      I_Contact( #s340_StWtOTSFrmTT_T1 )
      wire#w2
      Coil( #s340_StWtOTSFrmTT )
   END_RUNG
   RUNG wire#powerrail
      Contact( #s330_StWtL2S1Down_T1 )
   END_RUNG wire#w1
   RUNG wire#w2
      { S7_GenerateENO := "TRUE" } Move(in := 340, out1 => #StateNo)
   END_RUNG
   // the same network as SCL:
   #s340_StWtOTSFrmTT := (#s340_StWtOTSFrmTT OR #s330_StWtL2S1Down_T1) AND NOT #sStWtResetRel AND NOT #s340_StWtOTSFrmTT_T1;
   IF #s340_StWtOTSFrmTT THEN #StateNo := 340; END_IF;
END_REGION

REGION Network 94: Actions for STATE Num:340 StWtOTSFrmTT
   RUNG wire#powerrail
      Contact( #s340_StWtOTSFrmTT )
      Coil( #qRTRToTT )
   END_RUNG
   // the same network as SCL:
   #qRTRToTT := #s340_StWtOTSFrmTT;
END_REGION

REGION Network 95: Transition for STATE Num:350 StWtL2RecvingActive
   RUNG wire#powerrail
      Contact( #s350_StWtL2RecvingActive )
      I_Contact( #sStWtResetRel )
      Contact( #sSst )
      Contact( #iRecvAreaClear )
      Coil( #s350_StWtL2RecvingActive_T1 )
   END_RUNG
   // the same network as SCL:
   #s350_StWtL2RecvingActive_T1 := #s350_StWtL2RecvingActive AND NOT #sStWtResetRel AND #sSst AND #iRecvAreaClear;
END_REGION

REGION Network 96: STATE Num:350 StWtL2RecvingActive
   RUNG wire#powerrail
      Contact( #s350_StWtL2RecvingActive )
      wire#w1
      I_Contact( #sStWtResetRel )
      I_Contact( #s350_StWtL2RecvingActive_T1 )
      wire#w2
      Coil( #s350_StWtL2RecvingActive )
   END_RUNG
   RUNG wire#powerrail
      Contact( #s340_StWtOTSFrmTT_T1 )
   END_RUNG wire#w1
   RUNG wire#w2
      { S7_GenerateENO := "TRUE" } Move(in := 350, out1 => #StateNo)
   END_RUNG
   // the same network as SCL:
   #s350_StWtL2RecvingActive := (#s350_StWtL2RecvingActive OR #s340_StWtOTSFrmTT_T1) AND NOT #sStWtResetRel AND NOT #s350_StWtL2RecvingActive_T1;
   IF #s350_StWtL2RecvingActive THEN #StateNo := 350; END_IF;
END_REGION

REGION Network 97: Transition for STATE Num:360 StWtL2RcvDone
   RUNG wire#powerrail
      Contact( #s360_StWtL2RcvDone )
      I_Contact( #sStWtResetRel )
      Contact( #sSst )
      Contact( #iPalletAtL2 )
      Contact( #iReacvAreaClr )
      Coil( #s360_StWtL2RcvDone_T1 )
   END_RUNG
   // the same network as SCL:
   #s360_StWtL2RcvDone_T1 := #s360_StWtL2RcvDone AND NOT #sStWtResetRel AND #sSst AND #iPalletAtL2 AND #iReacvAreaClr;
END_REGION

REGION Network 98: STATE Num:360 StWtL2RcvDone
   RUNG wire#powerrail
      Contact( #s360_StWtL2RcvDone )
      wire#w1
      I_Contact( #sStWtResetRel )
      I_Contact( #s360_StWtL2RcvDone_T1 )
      wire#w2
      Coil( #s360_StWtL2RcvDone )
   END_RUNG
   RUNG wire#powerrail
      Contact( #s350_StWtL2RecvingActive_T1 )
   END_RUNG wire#w1
   RUNG wire#powerrail
      Contact( #s430_StNextRdyInTransit_3_T2 )
   END_RUNG wire#w1
   RUNG wire#w2
      { S7_GenerateENO := "TRUE" } Move(in := 360, out1 => #StateNo)
   END_RUNG
   // the same network as SCL:
   #s360_StWtL2RcvDone := (#s360_StWtL2RcvDone OR #s350_StWtL2RecvingActive_T1 OR #s430_StNextRdyInTransit_3_T2) AND NOT #sStWtResetRel AND NOT #s360_StWtL2RcvDone_T1;
   IF #s360_StWtL2RcvDone THEN #StateNo := 360; END_IF;
END_REGION

REGION Network 99: Transition for STATE Num:370 StChkPalAtTT
   RUNG wire#powerrail
      Contact( #s370_StChkPalAtTT )
      I_Contact( #sStWtResetRel )
      Contact( #sSst )
      wire#w1
      I_Contact( #ipalletPrsntAtTT )
      Coil( #s370_StChkPalAtTT_T1 )
   END_RUNG
   RUNG wire#w1
      I_Contact( #s370_StChkPalAtTT_T1 )
      Contact( #ipalletPrsntAtTT )
      Coil( #s370_StChkPalAtTT_T2 )
   END_RUNG
   RUNG wire#w1
      I_Contact( #s370_StChkPalAtTT_T1 )
      I_Contact( #s370_StChkPalAtTT_T2 )
      I_Contact( #ipalletPrsntAtTT )
      Coil( #s370_StChkPalAtTT_T3 )
   END_RUNG
   // the same network as SCL:
   #_w1 := #s370_StChkPalAtTT AND NOT #sStWtResetRel AND #sSst;
   #s370_StChkPalAtTT_T1 := #_w1 AND NOT #ipalletPrsntAtTT;
   #s370_StChkPalAtTT_T2 := #_w1 AND NOT #s370_StChkPalAtTT_T1 AND #ipalletPrsntAtTT;
   #s370_StChkPalAtTT_T3 := #_w1 AND NOT #s370_StChkPalAtTT_T1 AND NOT #s370_StChkPalAtTT_T2 AND NOT #ipalletPrsntAtTT;
END_REGION

REGION Network 100: STATE Num:370 StChkPalAtTT
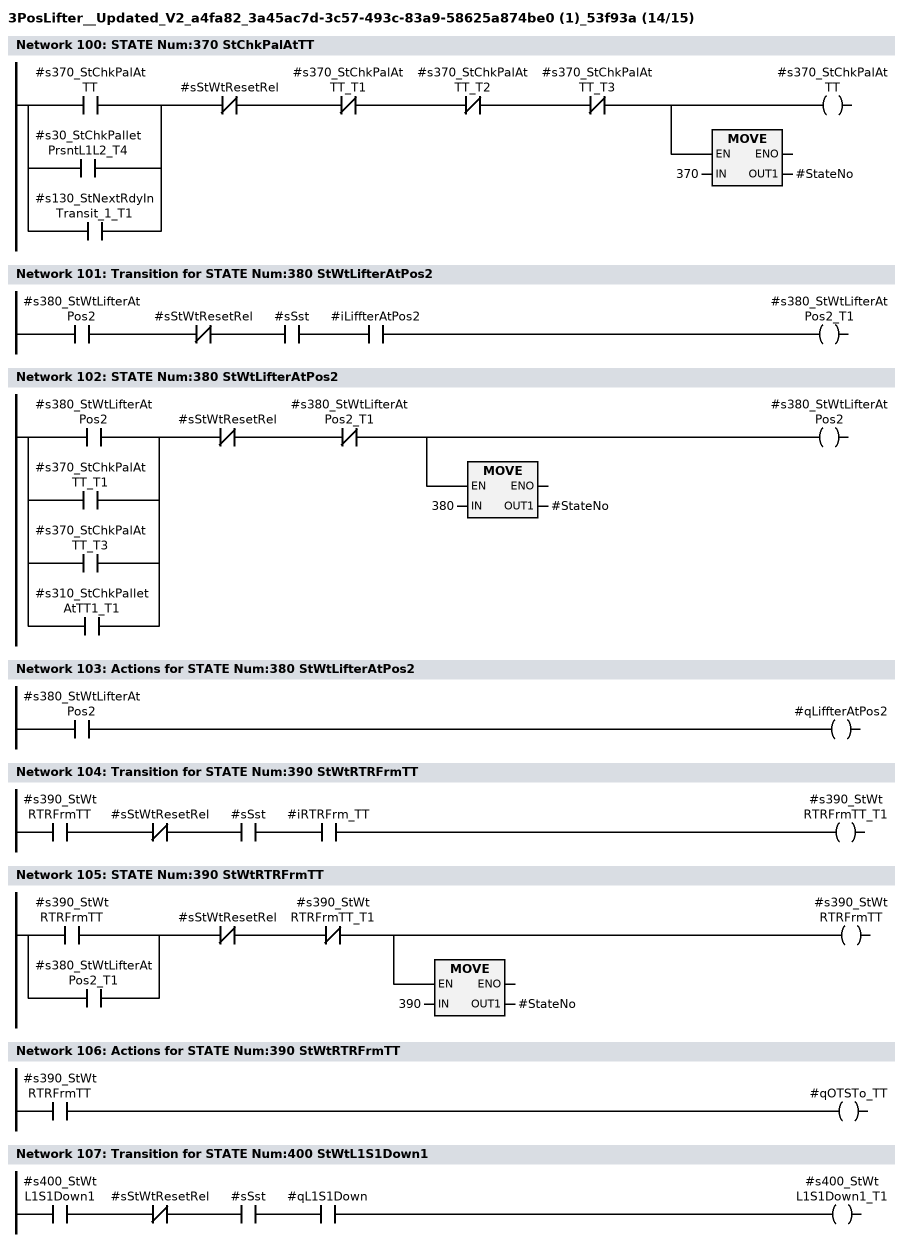
   RUNG wire#powerrail
      Contact( #s370_StChkPalAtTT )
      wire#w1
      I_Contact( #sStWtResetRel )
      I_Contact( #s370_StChkPalAtTT_T1 )
      I_Contact( #s370_StChkPalAtTT_T2 )
      I_Contact( #s370_StChkPalAtTT_T3 )
      wire#w2
      Coil( #s370_StChkPalAtTT )
   END_RUNG
   RUNG wire#powerrail
      Contact( #s30_StChkPalletPrsntL1L2_T4 )
   END_RUNG wire#w1
   RUNG wire#powerrail
      Contact( #s130_StNextRdyInTransit_1_T1 )
   END_RUNG wire#w1
   RUNG wire#w2
      { S7_GenerateENO := "TRUE" } Move(in := 370, out1 => #StateNo)
   END_RUNG
   // the same network as SCL:
   #s370_StChkPalAtTT := (#s370_StChkPalAtTT OR #s30_StChkPalletPrsntL1L2_T4 OR #s130_StNextRdyInTransit_1_T1) AND NOT #sStWtResetRel AND NOT #s370_StChkPalAtTT_T1 AND NOT #s370_StChkPalAtTT_T2 AND NOT #s370_StChkPalAtTT_T3;
   IF #s370_StChkPalAtTT THEN #StateNo := 370; END_IF;
END_REGION

REGION Network 101: Transition for STATE Num:380 StWtLifterAtPos2
   RUNG wire#powerrail
      Contact( #s380_StWtLifterAtPos2 )
      I_Contact( #sStWtResetRel )
      Contact( #sSst )
      Contact( #iLiffterAtPos2 )
      Coil( #s380_StWtLifterAtPos2_T1 )
   END_RUNG
   // the same network as SCL:
   #s380_StWtLifterAtPos2_T1 := #s380_StWtLifterAtPos2 AND NOT #sStWtResetRel AND #sSst AND #iLiffterAtPos2;
END_REGION

REGION Network 102: STATE Num:380 StWtLifterAtPos2
   RUNG wire#powerrail
      Contact( #s380_StWtLifterAtPos2 )
      wire#w1
      I_Contact( #sStWtResetRel )
      I_Contact( #s380_StWtLifterAtPos2_T1 )
      wire#w2
      Coil( #s380_StWtLifterAtPos2 )
   END_RUNG
   RUNG wire#powerrail
      Contact( #s370_StChkPalAtTT_T1 )
   END_RUNG wire#w1
   RUNG wire#powerrail
      Contact( #s370_StChkPalAtTT_T3 )
   END_RUNG wire#w1
   RUNG wire#powerrail
      Contact( #s310_StChkPalletAtTT1_T1 )
   END_RUNG wire#w1
   RUNG wire#w2
      { S7_GenerateENO := "TRUE" } Move(in := 380, out1 => #StateNo)
   END_RUNG
   // the same network as SCL:
   #s380_StWtLifterAtPos2 := (#s380_StWtLifterAtPos2 OR #s370_StChkPalAtTT_T1 OR #s370_StChkPalAtTT_T3 OR #s310_StChkPalletAtTT1_T1) AND NOT #sStWtResetRel AND NOT #s380_StWtLifterAtPos2_T1;
   IF #s380_StWtLifterAtPos2 THEN #StateNo := 380; END_IF;
END_REGION

REGION Network 103: Actions for STATE Num:380 StWtLifterAtPos2
   RUNG wire#powerrail
      Contact( #s380_StWtLifterAtPos2 )
      Coil( #qLiffterAtPos2 )
   END_RUNG
   // the same network as SCL:
   #qLiffterAtPos2 := #s380_StWtLifterAtPos2;
END_REGION

REGION Network 104: Transition for STATE Num:390 StWtRTRFrmTT
   RUNG wire#powerrail
      Contact( #s390_StWtRTRFrmTT )
      I_Contact( #sStWtResetRel )
      Contact( #sSst )
      Contact( #iRTRFrm_TT )
      Coil( #s390_StWtRTRFrmTT_T1 )
   END_RUNG
   // the same network as SCL:
   #s390_StWtRTRFrmTT_T1 := #s390_StWtRTRFrmTT AND NOT #sStWtResetRel AND #sSst AND #iRTRFrm_TT;
END_REGION

REGION Network 105: STATE Num:390 StWtRTRFrmTT
   RUNG wire#powerrail
      Contact( #s390_StWtRTRFrmTT )
      wire#w1
      I_Contact( #sStWtResetRel )
      I_Contact( #s390_StWtRTRFrmTT_T1 )
      wire#w2
      Coil( #s390_StWtRTRFrmTT )
   END_RUNG
   RUNG wire#powerrail
      Contact( #s380_StWtLifterAtPos2_T1 )
   END_RUNG wire#w1
   RUNG wire#w2
      { S7_GenerateENO := "TRUE" } Move(in := 390, out1 => #StateNo)
   END_RUNG
   // the same network as SCL:
   #s390_StWtRTRFrmTT := (#s390_StWtRTRFrmTT OR #s380_StWtLifterAtPos2_T1) AND NOT #sStWtResetRel AND NOT #s390_StWtRTRFrmTT_T1;
   IF #s390_StWtRTRFrmTT THEN #StateNo := 390; END_IF;
END_REGION

REGION Network 106: Actions for STATE Num:390 StWtRTRFrmTT
   RUNG wire#powerrail
      Contact( #s390_StWtRTRFrmTT )
      Coil( #qOTSTo_TT )
   END_RUNG
   // the same network as SCL:
   #qOTSTo_TT := #s390_StWtRTRFrmTT;
END_REGION

REGION Network 107: Transition for STATE Num:400 StWtL1S1Down1
   RUNG wire#powerrail
      Contact( #s400_StWtL1S1Down1 )
      I_Contact( #sStWtResetRel )
      Contact( #sSst )
      Contact( #qL1S1Down )
      Coil( #s400_StWtL1S1Down1_T1 )
   END_RUNG
   // the same network as SCL:
   #s400_StWtL1S1Down1_T1 := #s400_StWtL1S1Down1 AND NOT #sStWtResetRel AND #sSst AND #qL1S1Down;
END_REGION

REGION Network 108: STATE Num:400 StWtL1S1Down1
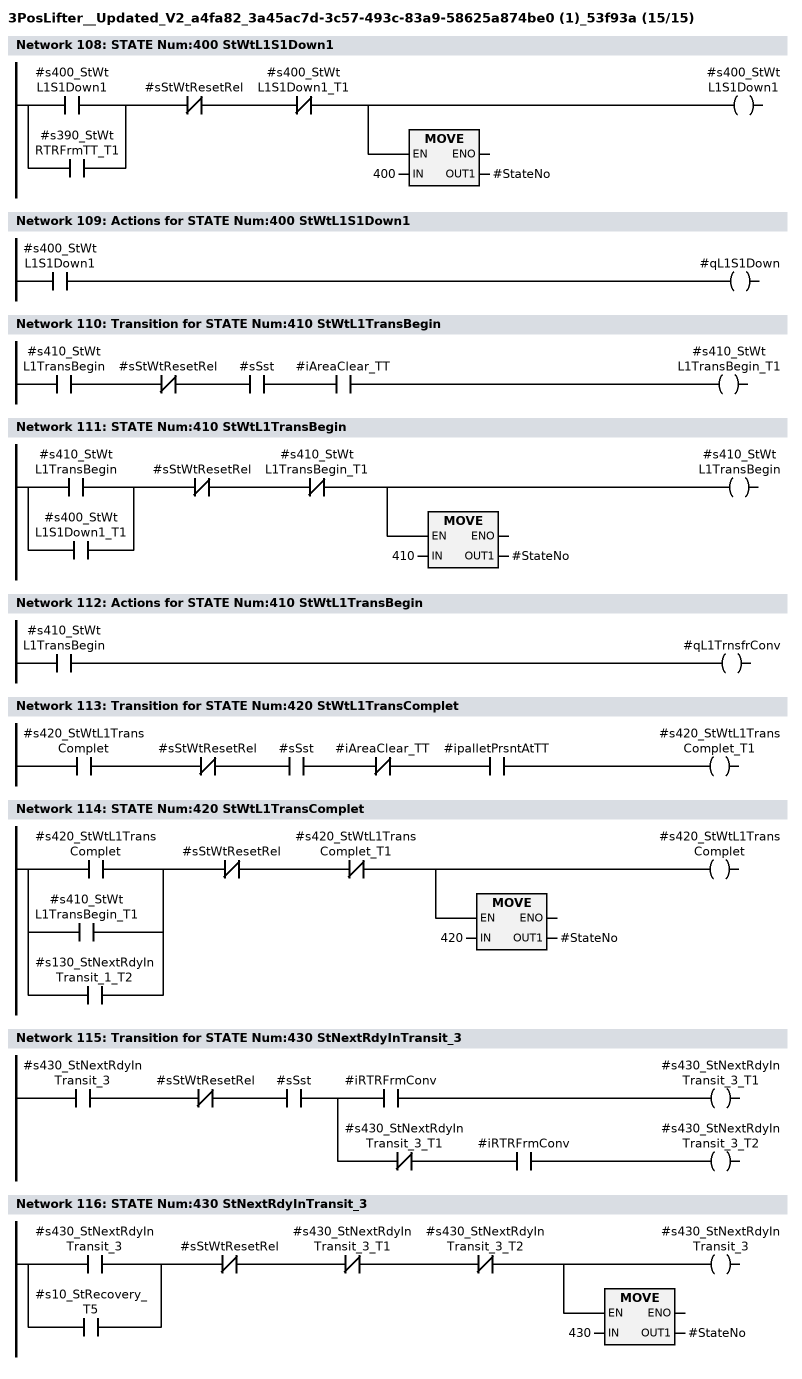
   RUNG wire#powerrail
      Contact( #s400_StWtL1S1Down1 )
      wire#w1
      I_Contact( #sStWtResetRel )
      I_Contact( #s400_StWtL1S1Down1_T1 )
      wire#w2
      Coil( #s400_StWtL1S1Down1 )
   END_RUNG
   RUNG wire#powerrail
      Contact( #s390_StWtRTRFrmTT_T1 )
   END_RUNG wire#w1
   RUNG wire#w2
      { S7_GenerateENO := "TRUE" } Move(in := 400, out1 => #StateNo)
   END_RUNG
   // the same network as SCL:
   #s400_StWtL1S1Down1 := (#s400_StWtL1S1Down1 OR #s390_StWtRTRFrmTT_T1) AND NOT #sStWtResetRel AND NOT #s400_StWtL1S1Down1_T1;
   IF #s400_StWtL1S1Down1 THEN #StateNo := 400; END_IF;
END_REGION

REGION Network 109: Actions for STATE Num:400 StWtL1S1Down1
   RUNG wire#powerrail
      Contact( #s400_StWtL1S1Down1 )
      Coil( #qL1S1Down )
   END_RUNG
   // the same network as SCL:
   #qL1S1Down := #s400_StWtL1S1Down1;
END_REGION

REGION Network 110: Transition for STATE Num:410 StWtL1TransBegin
   RUNG wire#powerrail
      Contact( #s410_StWtL1TransBegin )
      I_Contact( #sStWtResetRel )
      Contact( #sSst )
      Contact( #iAreaClear_TT )
      Coil( #s410_StWtL1TransBegin_T1 )
   END_RUNG
   // the same network as SCL:
   #s410_StWtL1TransBegin_T1 := #s410_StWtL1TransBegin AND NOT #sStWtResetRel AND #sSst AND #iAreaClear_TT;
END_REGION

REGION Network 111: STATE Num:410 StWtL1TransBegin
   RUNG wire#powerrail
      Contact( #s410_StWtL1TransBegin )
      wire#w1
      I_Contact( #sStWtResetRel )
      I_Contact( #s410_StWtL1TransBegin_T1 )
      wire#w2
      Coil( #s410_StWtL1TransBegin )
   END_RUNG
   RUNG wire#powerrail
      Contact( #s400_StWtL1S1Down1_T1 )
   END_RUNG wire#w1
   RUNG wire#w2
      { S7_GenerateENO := "TRUE" } Move(in := 410, out1 => #StateNo)
   END_RUNG
   // the same network as SCL:
   #s410_StWtL1TransBegin := (#s410_StWtL1TransBegin OR #s400_StWtL1S1Down1_T1) AND NOT #sStWtResetRel AND NOT #s410_StWtL1TransBegin_T1;
   IF #s410_StWtL1TransBegin THEN #StateNo := 410; END_IF;
END_REGION

REGION Network 112: Actions for STATE Num:410 StWtL1TransBegin
   RUNG wire#powerrail
      Contact( #s410_StWtL1TransBegin )
      Coil( #qL1TrnsfrConv )
   END_RUNG
   // the same network as SCL:
   #qL1TrnsfrConv := #s410_StWtL1TransBegin;
END_REGION

REGION Network 113: Transition for STATE Num:420 StWtL1TransComplet
   RUNG wire#powerrail
      Contact( #s420_StWtL1TransComplet )
      I_Contact( #sStWtResetRel )
      Contact( #sSst )
      I_Contact( #iAreaClear_TT )
      Contact( #ipalletPrsntAtTT )
      Coil( #s420_StWtL1TransComplet_T1 )
   END_RUNG
   // the same network as SCL:
   #s420_StWtL1TransComplet_T1 := #s420_StWtL1TransComplet AND NOT #sStWtResetRel AND #sSst AND NOT #iAreaClear_TT AND #ipalletPrsntAtTT;
END_REGION

REGION Network 114: STATE Num:420 StWtL1TransComplet
   RUNG wire#powerrail
      Contact( #s420_StWtL1TransComplet )
      wire#w1
      I_Contact( #sStWtResetRel )
      I_Contact( #s420_StWtL1TransComplet_T1 )
      wire#w2
      Coil( #s420_StWtL1TransComplet )
   END_RUNG
   RUNG wire#powerrail
      Contact( #s410_StWtL1TransBegin_T1 )
   END_RUNG wire#w1
   RUNG wire#powerrail
      Contact( #s130_StNextRdyInTransit_1_T2 )
   END_RUNG wire#w1
   RUNG wire#w2
      { S7_GenerateENO := "TRUE" } Move(in := 420, out1 => #StateNo)
   END_RUNG
   // the same network as SCL:
   #s420_StWtL1TransComplet := (#s420_StWtL1TransComplet OR #s410_StWtL1TransBegin_T1 OR #s130_StNextRdyInTransit_1_T2) AND NOT #sStWtResetRel AND NOT #s420_StWtL1TransComplet_T1;
   IF #s420_StWtL1TransComplet THEN #StateNo := 420; END_IF;
END_REGION

REGION Network 115: Transition for STATE Num:430 StNextRdyInTransit_3
   RUNG wire#powerrail
      Contact( #s430_StNextRdyInTransit_3 )
      I_Contact( #sStWtResetRel )
      Contact( #sSst )
      wire#w1
      Contact( #iRTRFrmConv )
      Coil( #s430_StNextRdyInTransit_3_T1 )
   END_RUNG
   RUNG wire#w1
      I_Contact( #s430_StNextRdyInTransit_3_T1 )
      Contact( #iRTRFrmConv )
      Coil( #s430_StNextRdyInTransit_3_T2 )
   END_RUNG
   // the same network as SCL:
   #_w1 := #s430_StNextRdyInTransit_3 AND NOT #sStWtResetRel AND #sSst;
   #s430_StNextRdyInTransit_3_T1 := #_w1 AND #iRTRFrmConv;
   #s430_StNextRdyInTransit_3_T2 := #_w1 AND NOT #s430_StNextRdyInTransit_3_T1 AND #iRTRFrmConv;
END_REGION

REGION Network 116: STATE Num:430 StNextRdyInTransit_3
   RUNG wire#powerrail
      Contact( #s430_StNextRdyInTransit_3 )
      wire#w1
      I_Contact( #sStWtResetRel )
      I_Contact( #s430_StNextRdyInTransit_3_T1 )
      I_Contact( #s430_StNextRdyInTransit_3_T2 )
      wire#w2
      Coil( #s430_StNextRdyInTransit_3 )
   END_RUNG
   RUNG wire#powerrail
      Contact( #s10_StRecovery_T5 )
   END_RUNG wire#w1
   RUNG wire#w2
      { S7_GenerateENO := "TRUE" } Move(in := 430, out1 => #StateNo)
   END_RUNG
   // the same network as SCL:
   #s430_StNextRdyInTransit_3 := (#s430_StNextRdyInTransit_3 OR #s10_StRecovery_T5) AND NOT #sStWtResetRel AND NOT #s430_StNextRdyInTransit_3_T1 AND NOT #s430_StNextRdyInTransit_3_T2;
   IF #s430_StNextRdyInTransit_3 THEN #StateNo := 430; END_IF;
END_REGION
END_FUNCTION_BLOCK

FUNCTION_BLOCK "3PosLifter__Updated_V2_a4fa82_3a45ac7d-3c57-493c-83a9-58625a874be0 (2) - Copy_22ffb1"   // FB1, STL
VERSION : 0.1
// stored: AutoNumber true, UDAEnableTagReadback false
   VAR_INPUT
      iAreaClearConv : Bool;
      iAreaClearTransL2 : Bool;
      iAreaClear_TT : Bool;
      iAutoRunning : Bool;
      iErrorAck : Bool;
      iL1PalletPrsnt : Bool;
      iL1S1Raise : Bool;
      iL1S2Down : Bool;
      iL1S2DownOver : Bool;
      iL2PalletPrsent : Bool;
      iL2S1Down : Bool;
      iL2S1Raise : Bool;
      iL2s2DownOver : Bool;
      iL2s2Raise : Bool;
      iLiffterAtPos1 : Bool;
      iLiffterAtPos2 : Bool;
      iLiffterAtPos3 : Bool;
      iLiffterAtPos4 : Bool;
      iLifterAt1 : Bool;
      iLifterAtPos1 : Bool;
      iLifterAtPos2 : Bool;
      iLifterAtPos3 : Bool;
      iLifterAtPos4 : Bool;
      iOTSFrmConv : Bool;
      iPalAtTT : Bool;
      iPalletAtL1 : Bool;
      iPalletAtL2 : Bool;
      iPalletAtTT : Bool;
      iPalletPrsntL1 : Bool;
      iRTRFrmConv : Bool;
      iRTRFrmTT : Bool;
      iRTRFrm_TT : Bool;
      iReacvAreaClr : Bool;
      iReceiveAreaClear : Bool;
      iReceiveAreaClrConv : Bool;
      iRecvAreaClear : Bool;
      iReset_fault : Bool;
      iRunOutActive : Bool;
      iRunOutCycle : Bool;
      iSstMode : Bool;
      iSstPB : Bool;
      iTransAreaClearConv : Bool;
      iTransAreaClr : Bool;
      ipalletPrsntAtTT : Bool;
   END_VAR
   VAR_OUTPUT
      qL1S1Down : Bool;
      qL1S1raise : Bool;
      qL1S2Down : Bool;
      qL1S2Raise : Bool;
      qL1TrnsfrConv : Bool;
      qL2S1raise : Bool;
      qL2S2Down : Bool;
      qL2S2Raise : Bool;
      qLiffterAtPos2 : Bool;
      qLifterAtPos1 : Bool;
      qLifterAtPos3 : Bool;
      qLifterAtPos4 : Bool;
      qLifterGotoPos1 : Bool;
      qOTSToNext : Bool;
      qOTSTo_TT : Bool;
      qOutput1 : Bool;
      qRTRToConv : Bool;
      qRTRToTT : Bool;
      qRTR_To_Conv : Bool;
   END_VAR
   VAR_IN_OUT
      IqRx_Frm_TT : Bool;
      iqRx_frm_Conv : Bool;
      iqTX_To_Conv : Bool;
      iqTX_To_TT : Bool;
      iqTx_To_ConvPos4 : Bool;
      iqTx_To_Rej : Bool;
   END_VAR
   VAR DB_SPECIFIC
      StateNo : Int;
      s190_sStWtL1RcvComplete_T1 : Bool;
      s200_sStWtForL1StprUp_T1 : Bool;
      s240_sStWtL2TransComplete_T1 : Bool;
      s250_sStWtDeforkDone : Bool;
      s250_sStWtDeforkDone_Cond1 : Bool;
      s250_sStWtDeforkDone_Cond2 : Bool;
      s250_sStWtDeforkDone_T1 : Bool;
      sInitialConvRun : Bool;
      sInitialConvRun_T1 : Bool;
      sOTSTimeout : Bool;
      sSeq1Over : Bool;
      sSeq2Over : Bool;
      sSst : Bool;
      sSstPulse : Bool;
      sSstRise : Bool;
      sStChkPalAtTT : Bool;
      sStChkPalAtTT_T1 : Bool;
      sStChkPalAtTT_T2 : Bool;
      sStChkPalAtTT_T3 : Bool;
      sStChkPalletAtTT : Bool;
      sStChkPalletAtTT1 : Bool;
      sStChkPalletAtTT1_T1 : Bool;
      sStChkPalletAtTT1_T2 : Bool;
      sStChkPalletAtTT_T1 : Bool;
      sStChkPalletAtTT_T2 : Bool;
      sStChkPalletPrsntL1L2 : Bool;
      sStChkPalletPrsntL1L2_T1 : Bool;
      sStChkPalletPrsntL1L2_T2 : Bool;
      sStChkPalletPrsntL1L2_T3 : Bool;
      sStChkPalletPrsntL1L2_T4 : Bool;
      sStChkRunOutActive1 : Bool;
      sStChkRunOutActive1_T1 : Bool;
      sStChkRunOutActive1_T2 : Bool;
      sStL1S2Down : Bool;
      sStL1S2DownOver : Bool;
      sStL1S2DownOver_T1 : Bool;
      sStL1S2Down_T1 : Bool;
      sStNextRdyInTransit : Bool;
      sStNextRdyInTransit_1 : Bool;
      sStNextRdyInTransit_1_T1 : Bool;
      sStNextRdyInTransit_1_T2 : Bool;
      sStNextRdyInTransit_3 : Bool;
      sStNextRdyInTransit_3_T1 : Bool;
      sStNextRdyInTransit_3_T2 : Bool;
      sStNextRdyInTransit_T1 : Bool;
      sStNextRdyInTransit_T2 : Bool;
      sStRecovery : Bool;
      sStRecovery_T1 : Bool;
      sStRecovery_T2 : Bool;
      sStRecovery_T3 : Bool;
      sStRecovery_T4 : Bool;
      sStRecovery_T5 : Bool;
      sStRecovery_T6 : Bool;
      sStRecovery_T7 : Bool;
      sStRecovery_T8 : Bool;
      sStRunOutActive : Bool;
      sStRunOutActive_T1 : Bool;
      sStRunOutActive_T2 : Bool;
      sStWtDeforkDone : Bool;
      sStWtDeforkDone_T1 : Bool;
      sStWtForFaultReset : Bool;
      sStWtForFaultReset_T1 : Bool;
      sStWtForL1L2StoprsUp : Bool;
      sStWtForL1L2StoprsUp_T1 : Bool;
      sStWtForL1StprUp : Bool;
      sStWtForL1StprUp_T1 : Bool;
      sStWtL1PalRcvDone : Bool;
      sStWtL1PalRcvDone_T1 : Bool;
      sStWtL1RcvComplete : Bool;
      sStWtL1RcvComplete_T1 : Bool;
      sStWtL1RecvBegin : Bool;
      sStWtL1RecvBegin_T1 : Bool;
      sStWtL1S1Down1 : Bool;
      sStWtL1S1Down1_T1 : Bool;
      sStWtL1S2DownOver : Bool;
      sStWtL1S2DownOver_T1 : Bool;
      sStWtL1TransBegin : Bool;
      sStWtL1TransBeginPos4 : Bool;
      sStWtL1TransBeginPos4_T1 : Bool;
      sStWtL1TransBegin_T1 : Bool;
      sStWtL1TransComplet : Bool;
      sStWtL1TransComplet_T1 : Bool;
      sStWtL2RcvDone : Bool;
      sStWtL2RcvDone_T1 : Bool;
      sStWtL2RecvingActive : Bool;
      sStWtL2RecvingActive_T1 : Bool;
      sStWtL2S1Down : Bool;
      sStWtL2S1Down_T1 : Bool;
      sStWtL2S2Down : Bool;
      sStWtL2S2Down_T1 : Bool;
      sStWtL2TranBegin : Bool;
      sStWtL2TranBegin_T1 : Bool;
      sStWtL2TransComplete : Bool;
      sStWtL2TransComplete_T1 : Bool;
      sStWtLifterAtPos1 : Bool;
      sStWtLifterAtPos1_T1 : Bool;
      sStWtLifterAtPos2 : Bool;
      sStWtLifterAtPos2_T1 : Bool;
      sStWtLifterAtPos3 : Bool;
      sStWtLifterAtPos3_T1 : Bool;
      sStWtLifterAtPos4 : Bool;
      sStWtLifterAtPos4_T1 : Bool;
      sStWtLifterAtPosn1 : Bool;
      sStWtLifterAtPosn1_T1 : Bool;
      sStWtOTSFrmConv : Bool;
      sStWtOTSFrmConv1 : Bool;
      sStWtOTSFrmConv1_T1 : Bool;
      sStWtOTSFrmConv1_T2 : Bool;
      sStWtOTSFrmConv_T1 : Bool;
      sStWtOTSFrmTT : Bool;
      sStWtOTSFrmTT_T1 : Bool;
      sStWtRTRFrmConvPos4 : Bool;
      sStWtRTRFrmConvPos4_T1 : Bool;
      sStWtRTRFrmTT : Bool;
      sStWtRTRFrmTT_T1 : Bool;
      sStWtRcvBegin : Bool;
      sStWtRcvBegin_T1 : Bool;
      sStWtResetRel : Bool;
      sStWtResetRel_T1 : Bool;
      sStWtTransDonePos4 : Bool;
      sStWtTransDonePos4_T1 : Bool;
   END_VAR
   VAR_TEMP
      tOne : Bool;
   END_VAR
BEGIN

NETWORK
TITLE = 
      O     #tOne;
      ON    #tOne;
      =     #tOne;

NETWORK
TITLE = Create Single Step Pulse bit
      A     #iSstPB;
      FP    #sSstRise;
      =     #sSstPulse;

NETWORK
TITLE = Create Single Step bit
      A     #iSstMode;
      A     #sSstPulse;
      ON    #iSstMode;
      =     #sSst;

NETWORK
TITLE = Transition for STATE Num:1 StWtResetRel
      A     #sStWtResetRel;
      AN    #sStWtResetRel;
      A     #sSst;
      A     #iAutoRunning;
      =     #sStWtResetRel_T1;

NETWORK
TITLE = STATE Num:1 StWtResetRel
      A(;
      O     #sStWtResetRel;
      ON    #iAutoRunning;
      );
      AN    #sStWtResetRel_T1;
      =     %L1.0;
      A     %L1.0;
      BLD   102;
      =     #sStWtResetRel;
      A     %L1.0;
      JNB   Label_1;
      L     1;
      T     #StateNo;
Label_1:NOP   0;

NETWORK
TITLE = Transition for STATE Num:10 StRecovery
      A     #sStRecovery;
      AN    #sStWtResetRel;
      A     #sSst;
      =     %L1.0;
      A     %L1.0;
      A(;
      O(;
      A     #iqTX_To_TT;
      AN    #iLifterAtPos2;
      );
      O(;
      A     #iqTX_To_Conv;
      AN    #iLifterAtPos1;
      );
      O(;
      A     #iqRx_frm_Conv;
      AN    #iLifterAtPos1;
      );
      O(;
      A     #IqRx_Frm_TT;
      AN    #iLifterAtPos3;
      );
      O(;
      A     #iqTx_To_Rej;
      AN    #iLifterAtPos4;
      );
      );
      =     #sStRecovery_T1;
      A     %L1.0;
      AN    #sStRecovery_T1;
      A     #iqTX_To_Conv;
      A     #iqRx_frm_Conv;
      A     #iLifterAtPos1;
      =     #sStRecovery_T2;
      A     %L1.0;
      AN    #sStRecovery_T1;
      AN    #sStRecovery_T2;
      A     #iqTX_To_TT;
      A     #iLifterAtPos2;
      =     #sStRecovery_T3;
      A     %L1.0;
      AN    #sStRecovery_T1;
      AN    #sStRecovery_T2;
      AN    #sStRecovery_T3;
      A     #iqTX_To_Conv;
      A     #iLifterAt1;
      =     #sStRecovery_T4;
      A     %L1.0;
      AN    #sStRecovery_T1;
      AN    #sStRecovery_T2;
      AN    #sStRecovery_T3;
      AN    #sStRecovery_T4;
      A     #iqTx_To_ConvPos4;
      A     #iLifterAtPos4;
      =     #sStRecovery_T5;
      A     %L1.0;
      AN    #sStRecovery_T1;
      AN    #sStRecovery_T2;
      AN    #sStRecovery_T3;
      AN    #sStRecovery_T4;
      AN    #sStRecovery_T5;
      A     #IqRx_Frm_TT;
      A     #iLifterAtPos3;
      =     #sStRecovery_T6;
      A     %L1.0;
      AN    #sStRecovery_T1;
      AN    #sStRecovery_T2;
      AN    #sStRecovery_T3;
      AN    #sStRecovery_T4;
      AN    #sStRecovery_T5;
      AN    #sStRecovery_T6;
      A     #iqRx_frm_Conv;
      A     #iLifterAtPos1;
      =     #sStRecovery_T7;
      A     %L1.0;
      AN    #sStRecovery_T1;
      AN    #sStRecovery_T2;
      AN    #sStRecovery_T3;
      AN    #sStRecovery_T4;
      AN    #sStRecovery_T5;
      AN    #sStRecovery_T6;
      AN    #sStRecovery_T7;
      AN    #iqTX_To_Conv;
      AN    #iqTX_To_TT;
      AN    #iqTx_To_ConvPos4;
      AN    #IqRx_Frm_TT;
      AN    #iqRx_frm_Conv;
      =     #sStRecovery_T8;

NETWORK
TITLE = STATE Num:10 StRecovery
      A(;
      O     #sStRecovery;
      O     #sInitialConvRun_T1;
      );
      AN    #sStWtResetRel;
      AN    #sStRecovery_T1;
      AN    #sStRecovery_T2;
      AN    #sStRecovery_T3;
      AN    #sStRecovery_T4;
      AN    #sStRecovery_T5;
      AN    #sStRecovery_T6;
      AN    #sStRecovery_T7;
      AN    #sStRecovery_T8;
      =     %L1.0;
      A     %L1.0;
      BLD   102;
      =     #sStRecovery;
      A     %L1.0;
      JNB   Label_10;
      L     10;
      T     #StateNo;
Label_10:NOP   0;

NETWORK
TITLE = Transition for STATE Num:15 StWtForFaultReset
      A     #sStWtForFaultReset;
      AN    #sStWtResetRel;
      A     #sSst;
      A     #iErrorAck;
      =     #sStWtForFaultReset_T1;

NETWORK
TITLE = STATE Num:15 StWtForFaultReset
      A(;
      O     #sStWtForFaultReset;
      O     #sStRecovery_T1;
      );
      AN    #sStWtResetRel;
      AN    #sStWtForFaultReset_T1;
      =     %L1.0;
      A     %L1.0;
      BLD   102;
      =     #sStWtForFaultReset;
      A     %L1.0;
      JNB   Label_15;
      L     15;
      T     #StateNo;
Label_15:NOP   0;

NETWORK
TITLE = Actions for STATE Num:15 StWtForFaultReset
      A     #sStWtForFaultReset;
      =     #qOutput1;

NETWORK
TITLE = Transition for STATE Num:20 StWtForL1L2StoprsUp
      A     #sStWtForL1L2StoprsUp;
      AN    #sStWtResetRel;
      A     #sSst;
      A     #iL1S1Raise;
      A     #iL1S1Raise;
      A     #iL2S1Raise;
      A     #iL2s2Raise;
      =     #sStWtForL1L2StoprsUp_T1;

NETWORK
TITLE = STATE Num:20 StWtForL1L2StoprsUp
      A(;
      O     #sStWtForL1L2StoprsUp;
      O     #sStRecovery_T8;
      O     #sStWtL1PalRcvDone_T1;
      O     #sStWtDeforkDone_T1;
      O     #sStWtTransDonePos4_T1;
      O     #sStWtL2RcvDone_T1;
      O     #sStWtL1TransComplet_T1;
      );
      AN    #sStWtResetRel;
      AN    #sStWtForL1L2StoprsUp_T1;
      =     %L1.0;
      A     %L1.0;
      BLD   102;
      =     #sStWtForL1L2StoprsUp;
      A     %L1.0;
      JNB   Label_20;
      L     20;
      T     #StateNo;
Label_20:NOP   0;

NETWORK
TITLE = Actions for STATE Num:20 StWtForL1L2StoprsUp
      A     #sStWtForL1L2StoprsUp;
      =     #qL1S1raise;
      =     #qL1S2Raise;
      =     #qL2S1raise;
      =     #qL2S2Raise;

NETWORK
TITLE = Transition for STATE Num:30 StChkPalletPrsntL1L2
      A     #sStChkPalletPrsntL1L2;
      AN    #sStWtResetRel;
      A     #sSst;
      =     %L1.0;
      A     %L1.0;
      AN    #iL1PalletPrsnt;
      AN    #iL2PalletPrsent;
      =     #sStChkPalletPrsntL1L2_T1;
      A     %L1.0;
      AN    #sStChkPalletPrsntL1L2_T1;
      AN    #iL1PalletPrsnt;
      A     #iL2PalletPrsent;
      =     #sStChkPalletPrsntL1L2_T2;
      A     %L1.0;
      AN    #sStChkPalletPrsntL1L2_T1;
      AN    #sStChkPalletPrsntL1L2_T2;
      A     #iL1PalletPrsnt;
      AN    #iL2PalletPrsent;
      =     #sStChkPalletPrsntL1L2_T3;
      A     %L1.0;
      AN    #sStChkPalletPrsntL1L2_T1;
      AN    #sStChkPalletPrsntL1L2_T2;
      AN    #sStChkPalletPrsntL1L2_T3;
      A     #iL1PalletPrsnt;
      A     #iL2PalletPrsent;
      =     #sStChkPalletPrsntL1L2_T4;

NETWORK
TITLE = STATE Num:30 StChkPalletPrsntL1L2
      A(;
      O     #sStChkPalletPrsntL1L2;
      O     #sStWtForL1L2StoprsUp_T1;
      );
      AN    #sStWtResetRel;
      AN    #sStChkPalletPrsntL1L2_T1;
      AN    #sStChkPalletPrsntL1L2_T2;
      AN    #sStChkPalletPrsntL1L2_T3;
      AN    #sStChkPalletPrsntL1L2_T4;
      =     %L1.0;
      A     %L1.0;
      BLD   102;
      =     #sStChkPalletPrsntL1L2;
      A     %L1.0;
      JNB   Label_30;
      L     30;
      T     #StateNo;
Label_30:NOP   0;

NETWORK
TITLE = Transition for STATE Num:40 StChkPalletAtTT
      A     #sStChkPalletAtTT;
      AN    #sStWtResetRel;
      A     #sSst;
      =     %L1.0;
      A     %L1.0;
      AN    #iPalletAtTT;
      =     #sStChkPalletAtTT_T1;
      A     %L1.0;
      AN    #sStChkPalletAtTT_T1;
      A     #ipalletPrsntAtTT;
      =     #sStChkPalletAtTT_T2;

NETWORK
TITLE = STATE Num:40 StChkPalletAtTT
      A(;
      O     #sStChkPalletAtTT;
      O     #sStChkPalletPrsntL1L2_T1;
      );
      AN    #sStWtResetRel;
      AN    #sStChkPalletAtTT_T1;
      AN    #sStChkPalletAtTT_T2;
      =     %L1.0;
      A     %L1.0;
      BLD   102;
      =     #sStChkPalletAtTT;
      A     %L1.0;
      JNB   Label_40;
      L     40;
      T     #StateNo;
Label_40:NOP   0;

NETWORK
TITLE = Transition for STATE Num:50 StWtLifterAtPos1
      A     #sStWtLifterAtPos1;
      AN    #sStWtResetRel;
      A     #sSst;
      A     #iLifterAtPos1;
      =     #sStWtLifterAtPos1_T1;

NETWORK
TITLE = STATE Num:50 StWtLifterAtPos1
      A(;
      O     #sStWtLifterAtPos1;
      O     #sStChkPalletAtTT_T1;
      O     #sStRunOutActive_T1;
      );
      AN    #sStWtResetRel;
      AN    #sStWtLifterAtPos1_T1;
      =     %L1.0;
      A     %L1.0;
      BLD   102;
      =     #sStWtLifterAtPos1;
      A     %L1.0;
      JNB   Label_50;
      L     50;
      T     #StateNo;
Label_50:NOP   0;

NETWORK
TITLE = Actions for STATE Num:50 StWtLifterAtPos1
      A     #sStWtLifterAtPos1;
      =     #qLifterGotoPos1;

NETWORK
TITLE = Transition for STATE Num:60 StWtL1S2DownOver
      A     #sStWtL1S2DownOver;
      AN    #sStWtResetRel;
      A     #sSst;
      A     #iL1S2DownOver;
      =     #sStWtL1S2DownOver_T1;

NETWORK
TITLE = STATE Num:60 StWtL1S2DownOver
      A(;
      O     #sStWtL1S2DownOver;
      O     #sStWtLifterAtPos1_T1;
      O     #sStRecovery_T7;
      );
      AN    #sStWtResetRel;
      AN    #sStWtL1S2DownOver_T1;
      =     %L1.0;
      A     %L1.0;
      BLD   102;
      =     #sStWtL1S2DownOver;
      A     %L1.0;
      JNB   Label_60;
      L     60;
      T     #StateNo;
Label_60:NOP   0;

NETWORK
TITLE = Actions for STATE Num:60 StWtL1S2DownOver
      A     #sStWtL1S2DownOver;
      =     #qL1S2Down;

NETWORK
TITLE = Transition for STATE Num:70 StWtOTSFrmConv
      A     #sStWtOTSFrmConv;
      AN    #sStWtResetRel;
      A     #sSst;
      A     #iOTSFrmConv;
      =     #sStWtOTSFrmConv_T1;

NETWORK
TITLE = STATE Num:70 StWtOTSFrmConv
      A(;
      O     #sStWtOTSFrmConv;
      O     #sStWtL1S2DownOver_T1;
      );
      AN    #sStWtResetRel;
      AN    #sStWtOTSFrmConv_T1;
      =     %L1.0;
      A     %L1.0;
      BLD   102;
      =     #sStWtOTSFrmConv;
      A     %L1.0;
      JNB   Label_70;
      L     70;
      T     #StateNo;
Label_70:NOP   0;

NETWORK
TITLE = Actions for STATE Num:70 StWtOTSFrmConv
      A     #sStWtOTSFrmConv;
      =     #qRTRToConv;

NETWORK
TITLE = Transition for STATE Num:80 StWtL1RecvBegin
      A     #sStWtL1RecvBegin;
      AN    #sStWtResetRel;
      A     #sSst;
      AN    #iReceiveAreaClear;
      =     #sStWtL1RecvBegin_T1;

NETWORK
TITLE = STATE Num:80 StWtL1RecvBegin
      A(;
      O     #sStWtL1RecvBegin;
      O     #sStWtOTSFrmConv_T1;
      );
      AN    #sStWtResetRel;
      AN    #sStWtL1RecvBegin_T1;
      =     %L1.0;
      A     %L1.0;
      BLD   102;
      =     #sStWtL1RecvBegin;
      A     %L1.0;
      JNB   Label_80;
      L     80;
      T     #StateNo;
Label_80:NOP   0;

NETWORK
TITLE = Transition for STATE Num:90 StWtL1PalRcvDone
      A     #sStWtL1PalRcvDone;
      AN    #sStWtResetRel;
      A     #sSst;
      A     #iL2PalletPrsent;
      A     #iReceiveAreaClrConv;
      =     #sStWtL1PalRcvDone_T1;

NETWORK
TITLE = STATE Num:90 StWtL1PalRcvDone
      A(;
      O     #sStWtL1PalRcvDone;
      O     #sStWtL1RecvBegin_T1;
      );
      AN    #sStWtResetRel;
      AN    #sStWtL1PalRcvDone_T1;
      =     %L1.0;
      A     %L1.0;
      BLD   102;
      =     #sStWtL1PalRcvDone;
      A     %L1.0;
      JNB   Label_90;
      L     90;
      T     #StateNo;
Label_90:NOP   0;

NETWORK
TITLE = Transition for STATE Num:100 StRunOutActive
      A     #sStRunOutActive;
      AN    #sStWtResetRel;
      A     #sSst;
      =     %L1.0;
      A     %L1.0;
      AN    #iRunOutCycle;
      =     #sStRunOutActive_T1;
      A     %L1.0;
      AN    #sStRunOutActive_T1;
      A     #iRunOutCycle;
      =     #sStRunOutActive_T2;

NETWORK
TITLE = STATE Num:100 StRunOutActive
      A(;
      O     #sStRunOutActive;
      O     #sStChkPalletAtTT_T2;
      );
      AN    #sStWtResetRel;
      AN    #sStRunOutActive_T1;
      AN    #sStRunOutActive_T2;
      =     %L1.0;
      A     %L1.0;
      BLD   102;
      =     #sStRunOutActive;
      A     %L1.0;
      JNB   Label_100;
      L     100;
      T     #StateNo;
Label_100:NOP   0;

NETWORK
TITLE = Transition for STATE Num:110 InitialConvRun
      A     #sInitialConvRun;
      AN    #sStWtResetRel;
      A     #sSst;
      A     #iLiffterAtPos1;
      A     #iLiffterAtPos2;
      A     #iLiffterAtPos3;
      A     #iLiffterAtPos4;
      =     #sInitialConvRun_T1;

NETWORK
TITLE = STATE Num:110 InitialConvRun
      A(;
      O     #sInitialConvRun;
//wrong transition variable removed
      );
      AN    #sStWtResetRel;
      AN    #sInitialConvRun_T1;
      =     %L1.0;
      A     %L1.0;
      BLD   102;
      =     #sInitialConvRun;
      A     %L1.0;
      JNB   Label_110;
      L     110;
      T     #StateNo;
Label_110:NOP   0;

NETWORK
TITLE = Transition for STATE Num:120 StNextRdyInTransit
      A     #sStNextRdyInTransit;
      AN    #sStWtResetRel;
      A     #sSst;
      =     %L1.0;
      A     %L1.0;
      A     #iRTRFrmConv;
      =     #sStNextRdyInTransit_T1;
      A     %L1.0;
      AN    #sStNextRdyInTransit_T1;
      AN    #iPalletAtL1;
      A     #iL1S1Raise;
      =     #sStNextRdyInTransit_T2;

NETWORK
TITLE = STATE Num:120 StNextRdyInTransit
      A(;
      O     #sStNextRdyInTransit;
      O     #sStRecovery_T4;
      O     #sStWtLifterAtPosn1_T1;
      );
      AN    #sStWtResetRel;
      AN    #sStNextRdyInTransit_T1;
      AN    #sStNextRdyInTransit_T2;
      =     %L1.0;
      A     %L1.0;
      BLD   102;
      =     #sStNextRdyInTransit;
      A     %L1.0;
      JNB   Label_120;
      L     120;
      T     #StateNo;
Label_120:NOP   0;

NETWORK
TITLE = Transition for STATE Num:130 StNextRdyInTransit_1
      A     #sStNextRdyInTransit_1;
      AN    #sStWtResetRel;
      A     #sSst;
      =     %L1.0;
      A     %L1.0;
      A     #iRTRFrmTT;
      =     #sStNextRdyInTransit_1_T1;
      A     %L1.0;
      AN    #sStNextRdyInTransit_1_T1;
      AN    #iPalletAtL1;
      A     #iL1S1Raise;
      =     #sStNextRdyInTransit_1_T2;

NETWORK
TITLE = STATE Num:130 StNextRdyInTransit_1
      A(;
      O     #sStNextRdyInTransit_1;
      O     #sStRecovery_T3;
      );
      AN    #sStWtResetRel;
      AN    #sStNextRdyInTransit_1_T1;
      AN    #sStNextRdyInTransit_1_T2;
      =     %L1.0;
      A     %L1.0;
      BLD   102;
      =     #sStNextRdyInTransit_1;
      A     %L1.0;
      JNB   Label_130;
      L     130;
      T     #StateNo;
Label_130:NOP   0;

NETWORK
TITLE = Transition for STATE Num:150 StWtLifterAtPosn1
      A     #sStWtLifterAtPosn1;
      AN    #sStWtResetRel;
      A     #sSst;
      A     #iLifterAtPos1;
      =     #sStWtLifterAtPosn1_T1;

NETWORK
TITLE = STATE Num:150 StWtLifterAtPosn1
      A(;
      O     #sStWtLifterAtPosn1;
      O     #sStChkPalletPrsntL1L2_T2;
      O     #sStRecovery_T2;
      O     #sStChkPalAtTT_T2;
      );
      AN    #sStWtResetRel;
      AN    #sStWtLifterAtPosn1_T1;
      =     %L1.0;
      A     %L1.0;
      BLD   102;
      =     #sStWtLifterAtPosn1;
      A     %L1.0;
      JNB   Label_150;
      L     150;
      T     #StateNo;
Label_150:NOP   0;

NETWORK
TITLE = Actions for STATE Num:150 StWtLifterAtPosn1
      A     #sStWtLifterAtPosn1;
      =     #qLifterAtPos1;

NETWORK
TITLE = Transition for STATE Num:160 StL1S2DownOver
      A     #sStL1S2DownOver;
      AN    #sStWtResetRel;
      A     #sSst;
      A     #iL1S2DownOver;
      =     #sStL1S2DownOver_T1;

NETWORK
TITLE = STATE Num:160 StL1S2DownOver
      A(;
      O     #sStL1S2DownOver;
      O     #sStWtLifterAtPosn1_T1;
      );
      AN    #sStWtResetRel;
      AN    #sStL1S2DownOver_T1;
      =     %L1.0;
      A     %L1.0;
      BLD   102;
      =     #sStL1S2DownOver;
      A     %L1.0;
      JNB   Label_160;
      L     160;
      T     #StateNo;
Label_160:NOP   0;

NETWORK
TITLE = Actions for STATE Num:160 StL1S2DownOver
      A     #sStL1S2DownOver;
      =     #qL1S2Down;

NETWORK
TITLE = Transition for STATE Num:170 StWtOTSFrmConv1
      A     #sStWtOTSFrmConv1;
      AN    #sStWtResetRel;
      A     #sSst;
      =     %L1.0;
      A     %L1.0;
      A     #iOTSFrmConv;
      =     #sStWtOTSFrmConv1_T1;
      A     %L1.0;
      AN    #sStWtOTSFrmConv1_T1;
      AN    #iOTSFrmConv;
      A     #sOTSTimeout;
      =     #sStWtOTSFrmConv1_T2;

NETWORK
TITLE = STATE Num:170 StWtOTSFrmConv1
      A(;
      O     #sStWtOTSFrmConv1;
      O     #sStL1S2DownOver_T1;
      );
      AN    #sStWtResetRel;
      AN    #sStWtOTSFrmConv1_T1;
      AN    #sStWtOTSFrmConv1_T2;
      =     %L1.0;
      A     %L1.0;
      BLD   102;
      =     #sStWtOTSFrmConv1;
      A     %L1.0;
      JNB   Label_170;
      L     170;
      T     #StateNo;
Label_170:NOP   0;

NETWORK
TITLE = Actions for STATE Num:170 StWtOTSFrmConv1
      A     #sStWtOTSFrmConv1;
      =     #qRTR_To_Conv;

NETWORK
TITLE = Transition for STATE Num:180 StWtRcvBegin
      A     #sStWtRcvBegin;
      AN    #sStWtResetRel;
      A     #sSst;
      AN    #iAreaClearConv;
      =     #sStWtRcvBegin_T1;

NETWORK
TITLE = STATE Num:180 StWtRcvBegin
      A(;
      O     #sStWtRcvBegin;
      O     #sStWtOTSFrmConv1_T1;
      );
      AN    #sStWtResetRel;
      AN    #sStWtRcvBegin_T1;
      =     %L1.0;
      A     %L1.0;
      BLD   102;
      =     #sStWtRcvBegin;
      A     %L1.0;
      JNB   Label_180;
      L     180;
      T     #StateNo;
Label_180:NOP   0;

NETWORK
TITLE = Transition for STATE Num:190 StWtL1RcvComplete
      A     #sStWtL1RcvComplete;
      AN    #sStWtResetRel;
      A     #sSst;
      A     #iPalletAtL1;
      A     #iAreaClearConv;
      =     #sStWtL1RcvComplete_T1;

NETWORK
TITLE = STATE Num:190 StWtL1RcvComplete
      A(;
      O     #sStWtL1RcvComplete;
      O     #sStWtRcvBegin_T1;
      );
      AN    #sStWtResetRel;
      AN    #sStWtL1RcvComplete_T1;
      =     %L1.0;
      A     %L1.0;
      BLD   102;
      =     #sStWtL1RcvComplete;
      A     %L1.0;
      JNB   Label_190;
      L     190;
      T     #StateNo;
Label_190:NOP   0;

NETWORK
TITLE = Transition for STATE Num:200 StWtForL1StprUp
      A     #sStWtForL1StprUp;
      AN    #sStWtResetRel;
      A     #sSst;
      A     #iL1S1Raise;
      A     #iL1S1Raise;
      =     #sStWtForL1StprUp_T1;

NETWORK
TITLE = STATE Num:200 StWtForL1StprUp
      A(;
      O     #sStWtForL1StprUp;
      O     #sStWtOTSFrmConv1_T2;
      );
      AN    #sStWtResetRel;
      AN    #sStWtForL1StprUp_T1;
      =     %L1.0;
      A     %L1.0;
      BLD   102;
      =     #sStWtForL1StprUp;
      A     %L1.0;
      JNB   Label_200;
      L     200;
      T     #StateNo;
Label_200:NOP   0;

NETWORK
TITLE = Actions for STATE Num:200 StWtForL1StprUp
      A     #sStWtForL1StprUp;
      =     #qL1S1raise;
      =     #qL1S2Raise;

NETWORK
TITLE = Transition for STATE Num:220 StWtL2S2Down
      A     #sStWtL2S2Down;
      AN    #sStWtResetRel;
      A     #sSst;
      A     #iL2s2DownOver;
      =     #sStWtL2S2Down_T1;

NETWORK
TITLE = STATE Num:220 StWtL2S2Down
      A(;
      O     #sStWtL2S2Down;
      O     #sStNextRdyInTransit_T1;
      );
      AN    #sStWtResetRel;
      AN    #sStWtL2S2Down_T1;
      =     %L1.0;
      A     %L1.0;
      BLD   102;
      =     #sStWtL2S2Down;
      A     %L1.0;
      JNB   Label_220;
      L     220;
      T     #StateNo;
Label_220:NOP   0;

NETWORK
TITLE = Actions for STATE Num:220 StWtL2S2Down
      A     #sStWtL2S2Down;
      =     #qL2S2Down;

NETWORK
TITLE = Transition for STATE Num:230 StWtL2TranBegin
      A     #sStWtL2TranBegin;
      AN    #sStWtResetRel;
      A     #sSst;
      AN    #iTransAreaClearConv;
      =     #sStWtL2TranBegin_T1;

NETWORK
TITLE = STATE Num:230 StWtL2TranBegin
      A(;
      O     #sStWtL2TranBegin;
      O     #sStWtL2S2Down_T1;
      );
      AN    #sStWtResetRel;
      AN    #sStWtL2TranBegin_T1;
      =     %L1.0;
      A     %L1.0;
      BLD   102;
      =     #sStWtL2TranBegin;
      A     %L1.0;
      JNB   Label_230;
      L     230;
      T     #StateNo;
Label_230:NOP   0;

NETWORK
TITLE = Transition for STATE Num:240 StWtL2TransComplete
      A     #sStWtL2TransComplete;
      AN    #sStWtResetRel;
      A     #sSst;
      AN    #iPalletAtL1;
      A     #iAreaClearTransL2;
      =     #sStWtL2TransComplete_T1;

NETWORK
TITLE = STATE Num:240 StWtL2TransComplete
      A(;
      O     #sStWtL2TransComplete;
      O     #sStWtL2TranBegin_T1;
      O     #sStNextRdyInTransit_T2;
      );
      AN    #sStWtResetRel;
      AN    #sStWtL2TransComplete_T1;
      =     %L1.0;
      A     %L1.0;
      BLD   102;
      =     #sStWtL2TransComplete;
      A     %L1.0;
      JNB   Label_240;
      L     240;
      T     #StateNo;
Label_240:NOP   0;

NETWORK
TITLE = Transition for STATE Num:250 Wait for event-1 to occur
      A     #s250_sStWtDeforkDone;
      AN    #sStWtResetRel;
      A     #sSst;
      A     #s250_sStWtDeforkDone_Cond1;  // Path 1 must be complete
      A     #s250_sStWtDeforkDone_Cond2;  // Path 2 must be complete
      AN    #sStWtL2TransComplete;  // condition expression
      AN    #sStWtL2TranBegin;  // condition expression
      AN    #sStWtForL1StprUp;  // condition expression
      A     #sSeq2Over;  // condition expression
      A     #sSeq1Over;  // condition expression
      =     #s250_sStWtDeforkDone_T1;


NETWORK
TITLE = Condition1 for STATE Num:250 Wait for event-1 to occur
      A(;
      O     #s190_sStWtL1RcvComplete_T1;  // Transition from state 190
      O     #s200_sStWtForL1StprUp_T1;  // Transition from state 200
      O     #s250_sStWtDeforkDone_Cond1;  // OR condition already set (self-latching)
      );
      AN    #sStWtResetRel;  // Reset signal must be inactive
      AN    #s250_sStWtDeforkDone_T1;  // Condition resets when state transitions out
      =     #s250_sStWtDeforkDone_Cond1;  // Set the condition flag for Path 1


NETWORK
TITLE = Condition2 for STATE Num:250 Wait for event-1 to occur
      A(;
      O     #s240_sStWtL2TransComplete_T1;  // Transition from state 240
      O     #s250_sStWtDeforkDone_Cond2;  // OR condition already set (self-latching)
      );
      AN    #sStWtResetRel;  // Reset signal must be inactive
      AN    #s250_sStWtDeforkDone_T1;  // Condition resets when state transitions out
      =     #s250_sStWtDeforkDone_Cond2;  // Set the condition flag for Path 2


NETWORK
TITLE = STATE Num:250 Wait for event-1 to occur
      A(;
      O     #s250_sStWtDeforkDone;  // state variable for state 250
      O     #s190_sStWtL1RcvComplete_T1;  // transition from state 190 in OR condition with state variable
      O     #s200_sStWtForL1StprUp_T1;  // transition from state 200 in OR condition with state variable
      O     #s240_sStWtL2TransComplete_T1;  // transition from state 240 in OR condition with state variable
      );
      AN    #sStWtResetRel;
      AN    #s250_sStWtDeforkDone_T1;
      =     %L1.0;
      A     %L1.0;
      BLD   102;
      =     #s250_sStWtDeforkDone;
      A     %L1.0;
      JNB   Label_250;
      L     250;
      T     #StateNo;
Label_250:NOP   0;


NETWORK
TITLE = Actions for STATE Num:250 StWtDeforkDone
      A     #sStWtDeforkDone;
      =     #qOutput1;

NETWORK
TITLE = Transition for STATE Num:260 StChkRunOutActive1
      A     #sStChkRunOutActive1;
      AN    #sStWtResetRel;
      A     #sSst;
      =     %L1.0;
      A     %L1.0;
      A     #iRunOutActive;
      =     #sStChkRunOutActive1_T1;
      A     %L1.0;
      AN    #sStChkRunOutActive1_T1;
      AN    #iRunOutActive;
      =     #sStChkRunOutActive1_T2;

NETWORK
TITLE = STATE Num:260 StChkRunOutActive1
      A(;
      O     #sStChkRunOutActive1;
      O     #sStChkPalletPrsntL1L2_T3;
      );
      AN    #sStWtResetRel;
      AN    #sStChkRunOutActive1_T1;
      AN    #sStChkRunOutActive1_T2;
      =     %L1.0;
      A     %L1.0;
      BLD   102;
      =     #sStChkRunOutActive1;
      A     %L1.0;
      JNB   Label_260;
      L     260;
      T     #StateNo;
Label_260:NOP   0;

NETWORK
TITLE = Transition for STATE Num:270 StWtLifterAtPos4
      A     #sStWtLifterAtPos4;
      AN    #sStWtResetRel;
      A     #sSst;
      A     #iLifterAtPos4;
      =     #sStWtLifterAtPos4_T1;

NETWORK
TITLE = STATE Num:270 StWtLifterAtPos4
      A(;
      O     #sStWtLifterAtPos4;
      O     #sStChkRunOutActive1_T1;
      );
      AN    #sStWtResetRel;
      AN    #sStWtLifterAtPos4_T1;
      =     %L1.0;
      A     %L1.0;
      BLD   102;
      =     #sStWtLifterAtPos4;
      A     %L1.0;
      JNB   Label_270;
      L     270;
      T     #StateNo;
Label_270:NOP   0;

NETWORK
TITLE = Actions for STATE Num:270 StWtLifterAtPos4
      A     #sStWtLifterAtPos4;
      =     #qLifterAtPos4;

NETWORK
TITLE = Transition for STATE Num:280 StWtRTRFrmConvPos4
      A     #sStWtRTRFrmConvPos4;
      AN    #sStWtResetRel;
      A     #sSst;
      A     #iRTRFrmConv;
      =     #sStWtRTRFrmConvPos4_T1;

NETWORK
TITLE = STATE Num:280 StWtRTRFrmConvPos4
      A(;
      O     #sStWtRTRFrmConvPos4;
      O     #sStWtLifterAtPos4_T1;
      O     #sStNextRdyInTransit_3_T1;
      );
      AN    #sStWtResetRel;
      AN    #sStWtRTRFrmConvPos4_T1;
      =     %L1.0;
      A     %L1.0;
      BLD   102;
      =     #sStWtRTRFrmConvPos4;
      A     %L1.0;
      JNB   Label_280;
      L     280;
      T     #StateNo;
Label_280:NOP   0;

NETWORK
TITLE = Actions for STATE Num:280 StWtRTRFrmConvPos4
      A     #sStWtRTRFrmConvPos4;
      =     #qOTSToNext;

NETWORK
TITLE = Transition for STATE Num:285 StL1S2Down
      A     #sStL1S2Down;
      AN    #sStWtResetRel;
      A     #sSst;
      A     #iL1S2Down;
      =     #sStL1S2Down_T1;

NETWORK
TITLE = STATE Num:285 StL1S2Down
      A(;
      O     #sStL1S2Down;
      O     #sStWtRTRFrmConvPos4_T1;
      );
      AN    #sStWtResetRel;
      AN    #sStL1S2Down_T1;
      =     %L1.0;
      A     %L1.0;
      BLD   102;
      =     #sStL1S2Down;
      A     %L1.0;
      JNB   Label_285;
      L     285;
      T     #StateNo;
Label_285:NOP   0;

NETWORK
TITLE = Actions for STATE Num:285 StL1S2Down
      A     #sStL1S2Down;
      =     #qL1S2Down;

NETWORK
TITLE = Transition for STATE Num:290 StWtL1TransBeginPos4
      A     #sStWtL1TransBeginPos4;
      AN    #sStWtResetRel;
      A     #sSst;
      AN    #iTransAreaClr;
      =     #sStWtL1TransBeginPos4_T1;

NETWORK
TITLE = STATE Num:290 StWtL1TransBeginPos4
      A(;
      O     #sStWtL1TransBeginPos4;
      O     #sStL1S2Down_T1;
      );
      AN    #sStWtResetRel;
      AN    #sStWtL1TransBeginPos4_T1;
      =     %L1.0;
      A     %L1.0;
      BLD   102;
      =     #sStWtL1TransBeginPos4;
      A     %L1.0;
      JNB   Label_290;
      L     290;
      T     #StateNo;
Label_290:NOP   0;

NETWORK
TITLE = Transition for STATE Num:300 StWtTransDonePos4
      A     #sStWtTransDonePos4;
      AN    #sStWtResetRel;
      A     #sSst;
      AN    #iPalletPrsntL1;
      A     #iTransAreaClr;
      =     #sStWtTransDonePos4_T1;

NETWORK
TITLE = STATE Num:300 StWtTransDonePos4
      A(;
      O     #sStWtTransDonePos4;
      O     #sStWtL1TransBeginPos4_T1;
      );
      AN    #sStWtResetRel;
      AN    #sStWtTransDonePos4_T1;
      =     %L1.0;
      A     %L1.0;
      BLD   102;
      =     #sStWtTransDonePos4;
      A     %L1.0;
      JNB   Label_300;
      L     300;
      T     #StateNo;
Label_300:NOP   0;

NETWORK
TITLE = Transition for STATE Num:310 StChkPalletAtTT1
      A     #sStChkPalletAtTT1;
      AN    #sStWtResetRel;
      A     #sSst;
      =     %L1.0;
      A     %L1.0;
      AN    #iPalAtTT;
      =     #sStChkPalletAtTT1_T1;
      A     %L1.0;
      AN    #sStChkPalletAtTT1_T1;
      AN    #iPalAtTT;
      =     #sStChkPalletAtTT1_T2;

NETWORK
TITLE = STATE Num:310 StChkPalletAtTT1
      A(;
      O     #sStChkPalletAtTT1;
      O     #sStChkRunOutActive1_T2;
      );
      AN    #sStWtResetRel;
      AN    #sStChkPalletAtTT1_T1;
      AN    #sStChkPalletAtTT1_T2;
      =     %L1.0;
      A     %L1.0;
      BLD   102;
      =     #sStChkPalletAtTT1;
      A     %L1.0;
      JNB   Label_310;
      L     310;
      T     #StateNo;
Label_310:NOP   0;

NETWORK
TITLE = Transition for STATE Num:320 StWtLifterAtPos3
      A     #sStWtLifterAtPos3;
      AN    #sStWtResetRel;
      A     #sSst;
      A     #iLifterAtPos3;
      =     #sStWtLifterAtPos3_T1;

NETWORK
TITLE = STATE Num:320 StWtLifterAtPos3
      A(;
      O     #sStWtLifterAtPos3;
      O     #sStChkPalletAtTT1_T2;
      O     #sStRunOutActive_T2;
      );
      AN    #sStWtResetRel;
      AN    #sStWtLifterAtPos3_T1;
      =     %L1.0;
      A     %L1.0;
      BLD   102;
      =     #sStWtLifterAtPos3;
      A     %L1.0;
      JNB   Label_320;
      L     320;
      T     #StateNo;
Label_320:NOP   0;

NETWORK
TITLE = Actions for STATE Num:320 StWtLifterAtPos3
      A     #sStWtLifterAtPos3;
      =     #qLifterAtPos3;

NETWORK
TITLE = Transition for STATE Num:330 StWtL2S1Down
      A     #sStWtL2S1Down;
      AN    #sStWtResetRel;
      A     #sSst;
      A     #iL2S1Down;
      =     #sStWtL2S1Down_T1;

NETWORK
TITLE = STATE Num:330 StWtL2S1Down
      A(;
      O     #sStWtL2S1Down;
      O     #sStWtLifterAtPos3_T1;
      O     #sStRecovery_T6;
      );
      AN    #sStWtResetRel;
      AN    #sStWtL2S1Down_T1;
      =     %L1.0;
      A     %L1.0;
      BLD   102;
      =     #sStWtL2S1Down;
      A     %L1.0;
      JNB   Label_330;
      L     330;
      T     #StateNo;
Label_330:NOP   0;

NETWORK
TITLE = Actions for STATE Num:330 StWtL2S1Down
      A     #sStWtL2S1Down;
      =     #qL1S1Down;

NETWORK
TITLE = Transition for STATE Num:340 StWtOTSFrmTT
      A     #sStWtOTSFrmTT;
      AN    #sStWtResetRel;
      A     #sSst;
      A     #iOTSFrmConv;
      =     #sStWtOTSFrmTT_T1;

NETWORK
TITLE = STATE Num:340 StWtOTSFrmTT
      A(;
      O     #sStWtOTSFrmTT;
      O     #sStWtL2S1Down_T1;
      );
      AN    #sStWtResetRel;
      AN    #sStWtOTSFrmTT_T1;
      =     %L1.0;
      A     %L1.0;
      BLD   102;
      =     #sStWtOTSFrmTT;
      A     %L1.0;
      JNB   Label_340;
      L     340;
      T     #StateNo;
Label_340:NOP   0;

NETWORK
TITLE = Actions for STATE Num:340 StWtOTSFrmTT
      A     #sStWtOTSFrmTT;
      =     #qRTRToTT;

NETWORK
TITLE = Transition for STATE Num:350 StWtL2RecvingActive
      A     #sStWtL2RecvingActive;
      AN    #sStWtResetRel;
      A     #sSst;
      A     #iRecvAreaClear;
      =     #sStWtL2RecvingActive_T1;

NETWORK
TITLE = STATE Num:350 StWtL2RecvingActive
      A(;
      O     #sStWtL2RecvingActive;
      O     #sStWtOTSFrmTT_T1;
      );
      AN    #sStWtResetRel;
      AN    #sStWtL2RecvingActive_T1;
      =     %L1.0;
      A     %L1.0;
      BLD   102;
      =     #sStWtL2RecvingActive;
      A     %L1.0;
      JNB   Label_350;
      L     350;
      T     #StateNo;
Label_350:NOP   0;

NETWORK
TITLE = Transition for STATE Num:360 StWtL2RcvDone
      A     #sStWtL2RcvDone;
      AN    #sStWtResetRel;
      A     #sSst;
      A     #iPalletAtL2;
      A     #iReacvAreaClr;
      =     #sStWtL2RcvDone_T1;

NETWORK
TITLE = STATE Num:360 StWtL2RcvDone
      A(;
      O     #sStWtL2RcvDone;
      O     #sStWtL2RecvingActive_T1;
      O     #sStNextRdyInTransit_3_T2;
      );
      AN    #sStWtResetRel;
      AN    #sStWtL2RcvDone_T1;
      =     %L1.0;
      A     %L1.0;
      BLD   102;
      =     #sStWtL2RcvDone;
      A     %L1.0;
      JNB   Label_360;
      L     360;
      T     #StateNo;
Label_360:NOP   0;

NETWORK
TITLE = Transition for STATE Num:370 StChkPalAtTT
      A     #sStChkPalAtTT;
      AN    #sStWtResetRel;
      A     #sSst;
      =     %L1.0;
      A     %L1.0;
      AN    #ipalletPrsntAtTT;
      =     #sStChkPalAtTT_T1;
      A     %L1.0;
      AN    #sStChkPalAtTT_T1;
      A     #ipalletPrsntAtTT;
      =     #sStChkPalAtTT_T2;
      A     %L1.0;
      AN    #sStChkPalAtTT_T1;
      AN    #sStChkPalAtTT_T2;
      AN    #ipalletPrsntAtTT;
      =     #sStChkPalAtTT_T3;

NETWORK
TITLE = STATE Num:370 StChkPalAtTT
      A(;
      O     #sStChkPalAtTT;
      O     #sStChkPalletPrsntL1L2_T4;
      O     #sStNextRdyInTransit_1_T1;
      );
      AN    #sStWtResetRel;
      AN    #sStChkPalAtTT_T1;
      AN    #sStChkPalAtTT_T2;
      AN    #sStChkPalAtTT_T3;
      =     %L1.0;
      A     %L1.0;
      BLD   102;
      =     #sStChkPalAtTT;
      A     %L1.0;
      JNB   Label_370;
      L     370;
      T     #StateNo;
Label_370:NOP   0;

NETWORK
TITLE = Transition for STATE Num:380 StWtLifterAtPos2
      A     #sStWtLifterAtPos2;
      AN    #sStWtResetRel;
      A     #sSst;
      A     #iLiffterAtPos2;
      =     #sStWtLifterAtPos2_T1;

NETWORK
TITLE = STATE Num:380 StWtLifterAtPos2
      A(;
      O     #sStWtLifterAtPos2;
      O     #sStChkPalAtTT_T1;
      O     #sStChkPalAtTT_T3;
      O     #sStChkPalletAtTT1_T1;
      );
      AN    #sStWtResetRel;
      AN    #sStWtLifterAtPos2_T1;
      =     %L1.0;
      A     %L1.0;
      BLD   102;
      =     #sStWtLifterAtPos2;
      A     %L1.0;
      JNB   Label_380;
      L     380;
      T     #StateNo;
Label_380:NOP   0;

NETWORK
TITLE = Actions for STATE Num:380 StWtLifterAtPos2
      A     #sStWtLifterAtPos2;
      =     #qLiffterAtPos2;

NETWORK
TITLE = Transition for STATE Num:390 StWtRTRFrmTT
      A     #sStWtRTRFrmTT;
      AN    #sStWtResetRel;
      A     #sSst;
      A     #iRTRFrm_TT;
      =     #sStWtRTRFrmTT_T1;

NETWORK
TITLE = STATE Num:390 StWtRTRFrmTT
      A(;
      O     #sStWtRTRFrmTT;
      O     #sStWtLifterAtPos2_T1;
      );
      AN    #sStWtResetRel;
      AN    #sStWtRTRFrmTT_T1;
      =     %L1.0;
      A     %L1.0;
      BLD   102;
      =     #sStWtRTRFrmTT;
      A     %L1.0;
      JNB   Label_390;
      L     390;
      T     #StateNo;
Label_390:NOP   0;

NETWORK
TITLE = Actions for STATE Num:390 StWtRTRFrmTT
      A     #sStWtRTRFrmTT;
      =     #qOTSTo_TT;

NETWORK
TITLE = Transition for STATE Num:400 StWtL1S1Down1
      A     #sStWtL1S1Down1;
      AN    #sStWtResetRel;
      A     #sSst;
      A     #qL1S1Down;
      =     #sStWtL1S1Down1_T1;

NETWORK
TITLE = STATE Num:400 StWtL1S1Down1
      A(;
      O     #sStWtL1S1Down1;
      O     #sStWtRTRFrmTT_T1;
      );
      AN    #sStWtResetRel;
      AN    #sStWtL1S1Down1_T1;
      =     %L1.0;
      A     %L1.0;
      BLD   102;
      =     #sStWtL1S1Down1;
      A     %L1.0;
      JNB   Label_400;
      L     400;
      T     #StateNo;
Label_400:NOP   0;

NETWORK
TITLE = Actions for STATE Num:400 StWtL1S1Down1
      A     #sStWtL1S1Down1;
      =     #qL1S1Down;

NETWORK
TITLE = Transition for STATE Num:410 StWtL1TransBegin
      A     #sStWtL1TransBegin;
      AN    #sStWtResetRel;
      A     #sSst;
      A     #iAreaClear_TT;
      =     #sStWtL1TransBegin_T1;

NETWORK
TITLE = STATE Num:410 StWtL1TransBegin
      A(;
      O     #sStWtL1TransBegin;
      O     #sStWtL1S1Down1_T1;
      );
      AN    #sStWtResetRel;
      AN    #sStWtL1TransBegin_T1;
      =     %L1.0;
      A     %L1.0;
      BLD   102;
      =     #sStWtL1TransBegin;
      A     %L1.0;
      JNB   Label_410;
      L     410;
      T     #StateNo;
Label_410:NOP   0;

NETWORK
TITLE = Actions for STATE Num:410 StWtL1TransBegin
      A     #sStWtL1TransBegin;
      =     #qL1TrnsfrConv;

NETWORK
TITLE = Transition for STATE Num:420 StWtL1TransComplet
      A     #sStWtL1TransComplet;
      AN    #sStWtResetRel;
      A     #sSst;
      AN    #iAreaClear_TT;
      A     #ipalletPrsntAtTT;
      =     #sStWtL1TransComplet_T1;

NETWORK
TITLE = STATE Num:420 StWtL1TransComplet
      A(;
      O     #sStWtL1TransComplet;
      O     #sStWtL1TransBegin_T1;
      O     #sStNextRdyInTransit_1_T2;
      );
      AN    #sStWtResetRel;
      AN    #sStWtL1TransComplet_T1;
      =     %L1.0;
      A     %L1.0;
      BLD   102;
      =     #sStWtL1TransComplet;
      A     %L1.0;
      JNB   Label_420;
      L     420;
      T     #StateNo;
Label_420:NOP   0;

NETWORK
TITLE = Transition for STATE Num:430 StNextRdyInTransit_3
      A     #sStNextRdyInTransit_3;
      AN    #sStWtResetRel;
      A     #sSst;
      =     %L1.0;
      A     %L1.0;
      A     #iRTRFrmConv;
      =     #sStNextRdyInTransit_3_T1;
      A     %L1.0;
      AN    #sStNextRdyInTransit_3_T1;
      A     #iRTRFrmConv;
      =     #sStNextRdyInTransit_3_T2;

NETWORK
TITLE = STATE Num:430 StNextRdyInTransit_3
      A(;
      O     #sStNextRdyInTransit_3;
      O     #sStRecovery_T5;
      );
      AN    #sStWtResetRel;
      AN    #sStNextRdyInTransit_3_T1;
      AN    #sStNextRdyInTransit_3_T2;
      =     %L1.0;
      A     %L1.0;
      BLD   102;
      =     #sStNextRdyInTransit_3;
      A     %L1.0;
      JNB   Label_430;
      L     430;
      T     #StateNo;
Label_430:NOP   0;
END_FUNCTION_BLOCK

